(* IEC 61131-3 sources: OpenUnit/plc/src, 8 files *)

(* ---- BMS.st ---- *)
(* BMS - Burner Management System (NFPA 85 style)
   Master fuel trip (MFT) with first-out cause, furnace purge (5 min) with permissives, gas
   fuel train (main gas trip valves / vent: double block and bleed), four burner elevation
   light-off sequences (igniter -> main flame proving -> in service, flame failure trips the
   elevation), light-off time limit, watchdog to the hardwired MFT relay in the field.
   The four elevations A..D are processed in a FOR loop over arrays 1..4: their field I/O is
   copied in at the top and out at the bottom.
   Naming: I_* field inputs, Q_* field outputs, P_<PEER>_* peer status, IO_* bridge signals. *)
PROGRAM BMS_MAIN
(*@IO*)
  VAR
    RT : FB_PLC_RUNTIME;
    T_AIRLOW : FB_TONS;
    T_LVLHH : FB_TONS;
    T_LVLLL : FB_TONS;
    T_FLAMELOSS : FB_TONS;
    T_FUELLOSS : FB_TONS;
    T_BFPLOSS : FB_TONS;
    T_HDRLL : FB_TONS;
    T_HDRHH : FB_TONS;
    T_SUPLOW : FB_TONS;
    dts : REAL;
    init : BOOL;
    (* process values *)
    idRun : BOOL;
    fdRun : BOOL;
    airPct : REAL;
    fp : REAL;
    lvl : REAL;
    hdr : REAL;
    sup : REAL;
    anyFlame : BOOL;
    anyBrnOpen : BOOL;
    nInService : DINT;
    bfpAny : BOOL;
    dehTripped : BOOL;
    dehTripPrev : BOOL;
    mgtvOpen : BOOL;
    (* MFT *)
    c : ARRAY[1..18] OF BOOL;   (* MFT conditions, by first-out cause number *)
    firstOut : DINT;
    mftOn : BOOL;
    cause : DINT;
    fuelWas : BOOL;
    lightoffT : REAL;
    lastFuel : REAL;
    (* purge *)
    ppFans : BOOL;
    ppAir : BOOL;
    ppFuelOff : BOOL;
    ppFurn : BOOL;
    ppDrum : BOOL;
    ppNoTrip : BOOL;
    ready : BOOL;
    purgeActive : BOOL;
    purgeT : REAL;
    purgeComplete : BOOL;
    (* gas train: 0 CLOSED, 1 OPENING, 2 OPEN, 3 TRIPPED *)
    trainState : DINT;
    trainT : REAL;
    trainPerm : BOOL;
    trainCmd : BOOL;
    trainOpen : BOOL;
    (* elevations: state 0 OFF, 1 STARTING, 2 IN SERVICE, 3 STOPPING, 4 FLAME FAIL *)
    x : INT;
    elevPerm : BOOL;
    eState : ARRAY[1..4] OF DINT;
    eT : ARRAY[1..4] OF REAL;
    eIgn : ARRAY[1..4] OF BOOL;
    eBrn : ARRAY[1..4] OF BOOL;
    eLossT : ARRAY[1..4] OF REAL;
    flame : ARRAY[1..4] OF BOOL;
    ignFlame : ARRAY[1..4] OF BOOL;
    brnOpen : ARRAY[1..4] OF BOOL;
    startPb : ARRAY[1..4] OF BOOL;
    stopPb : ARRAY[1..4] OF BOOL;
    fired : BOOL;
  END_VAR
  VAR CONSTANT
    AIR_MCR : REAL := 2247.0;       (* t/h *)
    PURGE_TIME : REAL := 300.0;     (* s *)
    LIGHTOFF_TIME : REAL := 900.0;  (* s *)
    S_OFF : DINT := 0;
    S_STARTING : DINT := 1;
    S_IN_SERVICE : DINT := 2;
    S_STOPPING : DINT := 3;
    S_FAIL : DINT := 4;
    TR_CLOSED : DINT := 0;
    TR_OPENING : DINT := 1;
    TR_OPEN : DINT := 2;
    TR_TRIPPED : DINT := 3;
  END_VAR

  (* ---------------------------------------------------------------- runtime services *)
  RT(SIM_MS := I_SIM_TIME_MS, IC_SEQ := IO_IC_SEQ, IC_ID := IO_IC_ID, IC_SNAP := IO_IC_SNAP, CYCLE_MS := 50.0,
     HEARTBEAT := HEARTBEAT, SCAN_COUNT := SCAN_COUNT, SCAN_MS := SCAN_MS, SIM_DT := SIM_DT,
     IC_APPLIED := IC_APPLIED, IC_ACK := IC_ACK);
  dts := RT.DTS;
  init := RT.IC_INIT;
  HEALTHY := IO_COMM_PLANT AND RT.READY;
  COMM_PLANT := IO_COMM_PLANT OR NOT RT.READY;   (* not reported before the bridge has initialised the PLC *)
  COMM_DEH := IO_COMM_DEH OR RT.GRACE OR NOT RT.READY;

  (* field I/O of the four elevations -> arrays *)
  flame[1] := I_FLAME_A; flame[2] := I_FLAME_B; flame[3] := I_FLAME_C; flame[4] := I_FLAME_D;
  ignFlame[1] := I_IGN_A_FLAME; ignFlame[2] := I_IGN_B_FLAME; ignFlame[3] := I_IGN_C_FLAME; ignFlame[4] := I_IGN_D_FLAME;
  brnOpen[1] := I_BRN_A_OPEN; brnOpen[2] := I_BRN_B_OPEN; brnOpen[3] := I_BRN_C_OPEN; brnOpen[4] := I_BRN_D_OPEN;
  startPb[1] := ELEV_A_START; startPb[2] := ELEV_B_START; startPb[3] := ELEV_C_START; startPb[4] := ELEV_D_START;
  stopPb[1] := ELEV_A_STOP; stopPb[2] := ELEV_B_STOP; stopPb[3] := ELEV_C_STOP; stopPb[4] := ELEV_D_STOP;

  (* ---------------------------------------------------------------- initial condition *)
  (* The firing state follows the plant: a fired boiler is on line with its burning elevations
     in service, otherwise the BMS starts tripped (cause 15, power-up) and needs a purge. *)
  IF init THEN
    fired := I_FLAME_A OR I_FLAME_B OR I_FLAME_C OR I_FLAME_D;
    purgeActive := FALSE;
    purgeT := 0.0;
    purgeComplete := FALSE;
    lightoffT := 0.0;
    dehTripPrev := FALSE;
    IF fired THEN
      mftOn := FALSE;
      cause := 0;
      fuelWas := TRUE;
      trainState := TR_OPEN;
    ELSE
      mftOn := TRUE;
      cause := 15;
      fuelWas := FALSE;
      trainState := TR_TRIPPED;
    END_IF;
    trainT := 0.0;
    FOR x := 1 TO 4 DO
      IF flame[x] THEN eState[x] := S_IN_SERVICE; ELSE eState[x] := S_OFF; END_IF;
      eT[x] := 60.0;
      eIgn[x] := FALSE;
      eBrn[x] := flame[x];
      eLossT[x] := 0.0;
    END_FOR;
    lastFuel := I_FUEL_HEAT;
  END_IF;

  IF RT.READY THEN
    idRun := I_ID_A_RUN OR I_ID_B_RUN;
    fdRun := I_FD_A_RUN OR I_FD_B_RUN;
    airPct := I_AIR_FLOW / AIR_MCR * 100.0;
    fp := MEDIAN3(I_FURN_PRESS_A, I_FURN_PRESS_B, I_FURN_PRESS_C);
    lvl := MEDIAN3(I_DRUM_LVL_A, I_DRUM_LVL_B, I_DRUM_LVL_C);
    hdr := I_GAS_HDR_PRESS;
    sup := I_GAS_SUPPLY_PRESS;
    anyFlame := FALSE;
    anyBrnOpen := FALSE;
    nInService := 0;
    FOR x := 1 TO 4 DO
      anyFlame := anyFlame OR flame[x];
      anyBrnOpen := anyBrnOpen OR brnOpen[x] OR eBrn[x];
      IF eState[x] = S_IN_SERVICE THEN nInService := nInService + 1; END_IF;
    END_FOR;
    bfpAny := I_BFP_A_RUN OR I_BFP_B_RUN OR I_BFP_C_RUN;
    dehTripped := IO_COMM_DEH AND P_DEH_TRIPPED;
    mgtvOpen := I_MGTV_OPEN;

    (* ---------------------------------------------------------------- MFT conditions *)
    T_AIRLOW(IN := airPct < 25.0, PT := 3.0, DTS := dts, INIT := init);
    T_LVLHH(IN := VOTE2OO3(I_DRUM_LVL_A > 250.0, I_DRUM_LVL_B > 250.0, I_DRUM_LVL_C > 250.0), PT := 3.0, DTS := dts, INIT := init);
    T_LVLLL(IN := VOTE2OO3(I_DRUM_LVL_A < -300.0, I_DRUM_LVL_B < -300.0, I_DRUM_LVL_C < -300.0), PT := 3.0, DTS := dts, INIT := init);
    T_FLAMELOSS(IN := anyBrnOpen AND NOT anyFlame, PT := 5.0, DTS := dts, INIT := init);
    T_FUELLOSS(IN := fuelWas AND NOT anyBrnOpen, PT := 2.0, DTS := dts, INIT := init);
    T_BFPLOSS(IN := fuelWas AND NOT bfpAny, PT := 10.0, DTS := dts, INIT := init);
    T_HDRLL(IN := nInService > 0 AND hdr < 120.0, PT := 2.0, DTS := dts, INIT := init);
    T_HDRHH(IN := mgtvOpen AND hdr > 4500.0, PT := 1.0, DTS := dts, INIT := init);
    T_SUPLOW(IN := mgtvOpen AND sup < 12.0, PT := 3.0, DTS := dts, INIT := init);
    c[1] := MFT_PB;                                                              (* manual *)
    c[2] := NOT idRun;                                                           (* both ID fans off *)
    c[3] := NOT fdRun;                                                           (* both FD fans off *)
    c[4] := T_AIRLOW.Q;                                                          (* air flow < 25 % *)
    c[5] := VOTE2OO3(I_FURN_PRESS_A > 20.0, I_FURN_PRESS_B > 20.0, I_FURN_PRESS_C > 20.0);    (* furnace HH *)
    c[6] := VOTE2OO3(I_FURN_PRESS_A < -25.0, I_FURN_PRESS_B < -25.0, I_FURN_PRESS_C < -25.0); (* furnace LL *)
    c[7] := T_LVLHH.Q;                                                           (* drum level HH *)
    c[8] := T_LVLLL.Q;                                                           (* drum level LL *)
    c[9] := T_FLAMELOSS.Q;                                                       (* loss of all flame *)
    c[10] := T_FUELLOSS.Q;                                                       (* loss of all fuel *)
    c[11] := dehTripped AND NOT dehTripPrev AND lastFuel > 0.4 * 1620.0;         (* turbine trip, firing > bypass *)
    c[12] := T_BFPLOSS.Q;                                                        (* all BFPs off *)
    c[13] := NOT mftOn AND NOT fuelWas AND lightoffT > LIGHTOFF_TIME;              (* light-off time expired *)
    c[14] := I_BMS_WD_FAIL;                                                      (* watchdog / field I/O *)
    c[15] := FALSE;                                                              (* power-up: set at initialisation *)
    c[16] := T_HDRLL.Q;                                                          (* gas header LL *)
    c[17] := T_HDRHH.Q;                                                          (* gas header HH *)
    c[18] := T_SUPLOW.Q;                                                         (* gas supply low *)
    dehTripPrev := dehTripped;
    lastFuel := I_FUEL_HEAT;
    IF NOT mftOn THEN
      lightoffT := lightoffT + dts;
      firstOut := FIRST_OUT(C1 := c[1], C2 := c[2], C3 := c[3], C4 := c[4], C5 := c[5], C6 := c[6], C7 := c[7], C8 := c[8], C9 := c[9],
                            C10 := c[10], C11 := c[11], C12 := c[12], C13 := c[13], C14 := c[14], C15 := c[15], C16 := c[16], C17 := c[17],
                            C18 := c[18]);
      IF firstOut > 0 THEN
        (* trip: first-out cause, purge lost, all elevations off *)
        mftOn := TRUE;
        cause := firstOut;
        purgeActive := FALSE;
        purgeT := 0.0;
        purgeComplete := FALSE;
        fuelWas := FALSE;
        FOR x := 1 TO 4 DO
          eState[x] := S_OFF;
          eIgn[x] := FALSE;
          eBrn[x] := FALSE;
        END_FOR;
      END_IF;
    END_IF;

    (* ---------------------------------------------------------------- purge *)
    ppFans := idRun AND fdRun;
    ppAir := airPct >= 25.0 AND airPct <= 40.0;
    ppFuelOff := I_MGTV_CLOSED;
    FOR x := 1 TO 4 DO
      ppFuelOff := ppFuelOff AND NOT brnOpen[x] AND NOT eIgn[x];
    END_FOR;
    ppFurn := ABS(fp) < 5.0;
    ppDrum := lvl > -250.0 AND lvl < 200.0;
    ppNoTrip := NOT (c[2] OR c[3] OR c[5] OR c[6] OR c[7] OR c[8] OR c[14]);
    PP_FANS := ppFans;
    PP_AIR := ppAir;
    PP_FUEL_OFF := ppFuelOff;
    PP_FURN := ppFurn;
    PP_DRUM := ppDrum;
    PP_NO_TRIP := ppNoTrip;
    ready := mftOn AND ppFans AND ppAir AND ppFuelOff AND ppFurn AND ppDrum AND ppNoTrip;
    IF PURGE_START AND ready AND NOT purgeComplete THEN
      purgeActive := TRUE;
      purgeT := 0.0;
      purgeComplete := FALSE;
    END_IF;
    IF purgeActive THEN
      IF NOT ready THEN
        purgeActive := FALSE;
      ELSE
        purgeT := purgeT + dts;
        IF purgeT >= PURGE_TIME THEN
          purgeActive := FALSE;
          purgeT := PURGE_TIME;
          purgeComplete := TRUE;
        END_IF;
      END_IF;
    END_IF;
    IF MFT_RESET AND mftOn AND purgeComplete AND ppNoTrip THEN
      mftOn := FALSE;
      cause := 0;
      purgeActive := FALSE;
      purgeT := 0.0;
      purgeComplete := FALSE;
      lightoffT := 0.0;
      fuelWas := FALSE;
      trainState := TR_CLOSED;
      trainT := 0.0;
    END_IF;

    (* ---------------------------------------------------------------- gas fuel train *)
    trainPerm := NOT mftOn AND sup > 16.0 AND I_MGTV_CLOSED;
    IF GAS_TRAIN_OPEN AND trainPerm AND trainState = TR_CLOSED THEN
      trainState := TR_OPENING;
      trainT := 0.0;
    END_IF;
    IF GAS_TRAIN_CLOSE AND nInService = 0 THEN
      trainState := TR_CLOSED;
      trainT := 0.0;
    END_IF;
    IF mftOn AND trainState <> TR_TRIPPED THEN
      trainState := TR_TRIPPED;
      trainT := 0.0;
    END_IF;
    IF trainState = TR_OPENING THEN
      trainT := trainT + dts;
      IF mgtvOpen THEN
        trainState := TR_OPEN;
      ELSIF trainT > 10.0 THEN
        trainState := TR_CLOSED;
        trainT := 0.0;
      END_IF;
    END_IF;
    trainCmd := trainState = TR_OPENING OR trainState = TR_OPEN;
    Q_MGTV_CMD := trainCmd;
    Q_GAS_VENT_CMD := NOT trainCmd;
    trainOpen := trainState = TR_OPEN AND mgtvOpen AND NOT I_GAS_VENT_OPEN;
    GAS_TRAIN_STATE := trainState;
    GAS_TRAIN_PERM := trainPerm;
    GAS_TRAIN_OPENED := trainOpen;

    (* ---------------------------------------------------------------- burner elevations *)
    elevPerm := NOT mftOn AND trainOpen AND airPct > 25.0 AND hdr > 150.0 AND hdr < 3000.0 AND ABS(fp) < 10.0;
    FOR x := 1 TO 4 DO
      IF startPb[x] AND elevPerm AND (eState[x] = S_OFF OR eState[x] = S_FAIL) THEN
        eState[x] := S_STARTING;
        eT[x] := 0.0;
      END_IF;
      IF stopPb[x] THEN
        IF eState[x] = S_STARTING OR eState[x] = S_IN_SERVICE THEN
          eState[x] := S_STOPPING;
          eT[x] := 0.0;
        ELSIF eState[x] = S_FAIL THEN
          eState[x] := S_OFF;
        END_IF;
      END_IF;
      eT[x] := eT[x] + dts;
      CASE eState[x] OF
        1: (* STARTING: igniter, then main burner valves once the igniter flame is proven *)
          eIgn[x] := TRUE;
          IF eT[x] > 6.0 AND NOT ignFlame[x] THEN
            eState[x] := S_FAIL; eIgn[x] := FALSE; eBrn[x] := FALSE; eT[x] := 0.0;   (* igniter flame not proven *)
          ELSIF ignFlame[x] THEN
            eBrn[x] := TRUE;
          END_IF;
          IF eState[x] = S_STARTING AND eBrn[x] AND flame[x] AND eT[x] > 5.0 THEN
            eState[x] := S_IN_SERVICE;
            eT[x] := 0.0;
          ELSIF eState[x] = S_STARTING AND eT[x] > 15.0 THEN
            eState[x] := S_FAIL; eIgn[x] := FALSE; eBrn[x] := FALSE; eT[x] := 0.0;   (* main flame not proven *)
          END_IF;
        2: (* IN SERVICE: igniter off after 10 s, 2 s loss of flame trips the elevation *)
          eBrn[x] := TRUE;
          eIgn[x] := eT[x] < 10.0;
          IF NOT flame[x] THEN eLossT[x] := MIN(2.0, eLossT[x] + dts); ELSE eLossT[x] := 0.0; END_IF;
          IF NOT flame[x] AND eLossT[x] >= 2.0 THEN
            eState[x] := S_FAIL; eIgn[x] := FALSE; eBrn[x] := FALSE; eT[x] := 0.0;   (* loss of flame *)
          END_IF;
        3: (* STOPPING *)
          eBrn[x] := FALSE;
          eIgn[x] := FALSE;
          IF eT[x] > 3.0 THEN eState[x] := S_OFF; END_IF;
      ELSE
        eBrn[x] := FALSE;
        eIgn[x] := FALSE;
      END_CASE;
      IF eState[x] <> S_IN_SERVICE THEN eLossT[x] := 0.0; END_IF;
      IF mftOn THEN
        eBrn[x] := FALSE;
        eIgn[x] := FALSE;
        IF eState[x] <> S_FAIL THEN eState[x] := S_OFF; END_IF;
      END_IF;
    END_FOR;
    nInService := 0;
    FOR x := 1 TO 4 DO
      IF eState[x] = S_IN_SERVICE THEN nInService := nInService + 1; END_IF;
    END_FOR;
    IF nInService > 0 THEN fuelWas := TRUE; END_IF;

    (* arrays -> field outputs and faceplate status *)
    Q_IGN_A_CMD := eIgn[1]; Q_IGN_B_CMD := eIgn[2]; Q_IGN_C_CMD := eIgn[3]; Q_IGN_D_CMD := eIgn[4];
    Q_BRN_A_CMD := eBrn[1]; Q_BRN_B_CMD := eBrn[2]; Q_BRN_C_CMD := eBrn[3]; Q_BRN_D_CMD := eBrn[4];
    ELEV_A_STATE := eState[1]; ELEV_B_STATE := eState[2]; ELEV_C_STATE := eState[3]; ELEV_D_STATE := eState[4];
    ELEV_A_INSERV := eState[1] = S_IN_SERVICE; ELEV_B_INSERV := eState[2] = S_IN_SERVICE;
    ELEV_C_INSERV := eState[3] = S_IN_SERVICE; ELEV_D_INSERV := eState[4] = S_IN_SERVICE;
    ELEV_A_FAIL := eState[1] = S_FAIL; ELEV_B_FAIL := eState[2] = S_FAIL;
    ELEV_C_FAIL := eState[3] = S_FAIL; ELEV_D_FAIL := eState[4] = S_FAIL;
    ELEV_A_PERM := elevPerm; ELEV_B_PERM := elevPerm; ELEV_C_PERM := elevPerm; ELEV_D_PERM := elevPerm;

    (* ---------------------------------------------------------------- outputs & status *)
    Q_MFT_TRIP := mftOn;
    MFT := mftOn;
    MFT_CAUSE := cause;
    PURGE_READY := ready;
    PURGE_ACTIVE := purgeActive;
    PURGE_COMPLETE := purgeComplete;
    IF purgeComplete THEN PURGE_REMAIN := 0.0; ELSE PURGE_REMAIN := PURGE_TIME - purgeT; END_IF;
    IF mftOn OR fuelWas THEN LIGHTOFF_REMAIN := 0.0; ELSE LIGHTOFF_REMAIN := MAX(0.0, LIGHTOFF_TIME - lightoffT); END_IF;
    FUEL_IN_SERVICE := nInService > 0;
    ELEV_INSERV := nInService;
    IF anyFlame THEN FIREBALL := MIN(100.0, I_FUEL_HEAT / 1620.0 * 110.0); ELSE FIREBALL := 0.0; END_IF;
  END_IF;

  (* watchdog to the hardwired MFT relay: the field trips the boiler if this stops changing *)
  Q_BMS_WD := HEARTBEAT;

  (* operator pulses are consumed in the scan they arrive *)
  MFT_PB := FALSE;
  PURGE_START := FALSE;
  MFT_RESET := FALSE;
  GAS_TRAIN_OPEN := FALSE;
  GAS_TRAIN_CLOSE := FALSE;
  ELEV_A_START := FALSE; ELEV_B_START := FALSE; ELEV_C_START := FALSE; ELEV_D_START := FALSE;
  ELEV_A_STOP := FALSE; ELEV_B_STOP := FALSE; ELEV_C_STOP := FALSE; ELEV_D_STOP := FALSE;
END_PROGRAM

(* ---- BOP.st ---- *)
(* BOP - Balance of Plant / Turbine Auxiliaries
   Circulating water, condenser vacuum, condensate pumps, lube oil / jacking oil / turning
   gear, gland steam, vacuum breaker, hotwell level (condenser make-up).
   Naming: I_* field inputs, Q_* field outputs, P_<PEER>_* peer status, IO_* bridge signals;
   all other located variables are this controller's own Modbus registers (HMI faceplates). *)
PROGRAM BOP_MAIN
(*@IO*)
  VAR
    RT : FB_PLC_RUNTIME;
    CWP_A : FB_MOTOR;
    CWP_B : FB_MOTOR;
    VP_A : FB_MOTOR;
    VP_B : FB_MOTOR;
    CEP_A : FB_MOTOR;
    CEP_B : FB_MOTOR;
    AOP : FB_MOTOR;
    EOP : FB_MOTOR;
    JOP : FB_MOTOR;
    TG : FB_MOTOR;
    GLAND : FB_ONOFF;
    VB : FB_ONOFF;
    HW_DUMP : FB_ONOFF;
    LIC_HW : FB_LOOP;
    CEP_LOWP_TMR : FB_TONS;
    dts : REAL;
    init : BOOL;
    speed : REAL;
    condP : REAL;
    loP : REAL;
    hwLvl : REAL;
    vacPoor : BOOL;
    cepPermit : BOOL;
    cepLowP : BOOL;
    tgPermit : BOOL;
    dehTripped : BOOL;
    tripCwpA : BOOL;
    tripCwpB : BOOL;
    tripVpA : BOOL;
    tripVpB : BOOL;
    tripCepA : BOOL;
    tripCepB : BOOL;
  END_VAR

  (* ---------------------------------------------------------------- runtime services *)
  RT(SIM_MS := I_SIM_TIME_MS, IC_SEQ := IO_IC_SEQ, IC_ID := IO_IC_ID, IC_SNAP := IO_IC_SNAP, CYCLE_MS := 50.0,
     HEARTBEAT := HEARTBEAT, SCAN_COUNT := SCAN_COUNT, SCAN_MS := SCAN_MS, SIM_DT := SIM_DT,
     IC_APPLIED := IC_APPLIED, IC_ACK := IC_ACK);
  dts := RT.DTS;
  init := RT.IC_INIT;
  HEALTHY := IO_COMM_PLANT AND RT.READY;
  COMM_PLANT := IO_COMM_PLANT OR NOT RT.READY;   (* not reported before the bridge has initialised the PLC *)
  COMM_DEH := IO_COMM_DEH OR RT.GRACE OR NOT RT.READY;

  (* ---------------------------------------------------------------- built-in initial condition *)
  IF RT.IC_BUILTIN THEN
    CWP_A_MODE := 1; CWP_B_MODE := 1; VP_A_MODE := 1; VP_B_MODE := 1; CEP_A_MODE := 1; CEP_B_MODE := 1;
    AOP_MODE := 1; EOP_MODE := 1; JOP_MODE := 1; TG_MODE := 1;
    HW_DUMP_MODE := 1;
    LIC_HW_OUT := I_MAKEUP_FB;
    IF IO_IC_ID >= 2 THEN
      LIC_HW_MODE := 1;
    ELSE
      LIC_HW_MODE := 0;
    END_IF;
  END_IF;

  IF RT.READY THEN
    speed := MEDIAN3(I_SPEED_A, I_SPEED_B, I_SPEED_C);
    condP := I_COND_PRESS;
    loP := I_LO_PRESS;
    hwLvl := I_HW_LVL;

    (* Standby pumps start on the latched trip of the duty pump (cleared by the operator's STOP) *)
    tripCwpA := I_CWP_A_TRIP OR (CWP_A.LATCHED AND NOT init);
    tripCwpB := I_CWP_B_TRIP OR (CWP_B.LATCHED AND NOT init);
    tripVpA := I_VP_A_TRIP OR (VP_A.LATCHED AND NOT init);
    tripVpB := I_VP_B_TRIP OR (VP_B.LATCHED AND NOT init);
    tripCepA := I_CEP_A_TRIP OR (CEP_A.LATCHED AND NOT init);
    tripCepB := I_CEP_B_TRIP OR (CEP_B.LATCHED AND NOT init);

    (* ---- circulating water: the standby pump starts when the duty pump trips *)
    CWP_A(RUN_FB := I_CWP_A_RUN, TRIP_FB := I_CWP_A_TRIP, AUTO_START := tripCwpB, SYNC := init,
          START := CWP_A_START, STOP := CWP_A_STOP, MODE := CWP_A_MODE, CMD := Q_CWP_A_CMD,
          RUN := CWP_A_RUN, TRIP := CWP_A_TRIP, PERM := CWP_A_PERM, ILK_T := CWP_A_ILK);
    CWP_B(RUN_FB := I_CWP_B_RUN, TRIP_FB := I_CWP_B_TRIP, AUTO_START := tripCwpA, SYNC := init,
          START := CWP_B_START, STOP := CWP_B_STOP, MODE := CWP_B_MODE, CMD := Q_CWP_B_CMD,
          RUN := CWP_B_RUN, TRIP := CWP_B_TRIP, PERM := CWP_B_PERM, ILK_T := CWP_B_ILK);

    (* ---- vacuum pumps: standby starts on partner trip or poor vacuum *)
    vacPoor := condP > 150.0 AND I_GLAND_ON;
    VP_A(RUN_FB := I_VP_A_RUN, TRIP_FB := I_VP_A_TRIP, AUTO_START := tripVpB OR (vacPoor AND I_VP_B_RUN), SYNC := init,
         START := VP_A_START, STOP := VP_A_STOP, MODE := VP_A_MODE, CMD := Q_VP_A_CMD,
         RUN := VP_A_RUN, TRIP := VP_A_TRIP, PERM := VP_A_PERM, ILK_T := VP_A_ILK);
    VP_B(RUN_FB := I_VP_B_RUN, TRIP_FB := I_VP_B_TRIP, AUTO_START := tripVpA OR (vacPoor AND I_VP_A_RUN), SYNC := init,
         START := VP_B_START, STOP := VP_B_STOP, MODE := VP_B_MODE, CMD := Q_VP_B_CMD,
         RUN := VP_B_RUN, TRIP := VP_B_TRIP, PERM := VP_B_PERM, ILK_T := VP_B_ILK);

    (* ---- condensate pumps: need hotwell level; standby starts on trip or low discharge pressure *)
    cepPermit := hwLvl > 300.0;
    CEP_LOWP_TMR(IN := I_CEP_PRESS < 12.0 AND (I_CEP_A_RUN OR I_CEP_B_RUN), PT := 5.0, DTS := dts, INIT := init);
    cepLowP := CEP_LOWP_TMR.Q;
    CEP_A(RUN_FB := I_CEP_A_RUN, TRIP_FB := I_CEP_A_TRIP, PERMIT := cepPermit, AUTO_START := tripCepB OR (cepLowP AND I_CEP_B_RUN), SYNC := init,
          START := CEP_A_START, STOP := CEP_A_STOP, MODE := CEP_A_MODE, CMD := Q_CEP_A_CMD,
          RUN := CEP_A_RUN, TRIP := CEP_A_TRIP, PERM := CEP_A_PERM, ILK_T := CEP_A_ILK);
    CEP_B(RUN_FB := I_CEP_B_RUN, TRIP_FB := I_CEP_B_TRIP, PERMIT := cepPermit, AUTO_START := tripCepA OR (cepLowP AND I_CEP_A_RUN), SYNC := init,
          START := CEP_B_START, STOP := CEP_B_STOP, MODE := CEP_B_MODE, CMD := Q_CEP_B_CMD,
          RUN := CEP_B_RUN, TRIP := CEP_B_TRIP, PERM := CEP_B_PERM, ILK_T := CEP_B_ILK);

    (* ---- lube oil, jacking oil, turning gear *)
    AOP(RUN_FB := I_AOP_RUN, TRIP_FB := I_AOP_TRIP, AUTO_START := loP < 1.0, SYNC := init,
        START := AOP_START, STOP := AOP_STOP, MODE := AOP_MODE, CMD := Q_AOP_CMD,
        RUN := AOP_RUN, TRIP := AOP_TRIP, PERM := AOP_PERM, ILK_T := AOP_ILK);
    EOP(RUN_FB := I_EOP_RUN, TRIP_FB := I_EOP_TRIP, AUTO_START := loP < 0.7, SYNC := init,
        START := EOP_START, STOP := EOP_STOP, MODE := EOP_MODE, CMD := Q_EOP_CMD,
        RUN := EOP_RUN, TRIP := EOP_TRIP, PERM := EOP_PERM, ILK_T := EOP_ILK);
    JOP(RUN_FB := I_JOP_RUN, TRIP_FB := I_JOP_TRIP, AUTO_START := speed < 600.0 AND loP > 0.5, AUTO_STOP := speed > 700.0, SYNC := init,
        START := JOP_START, STOP := JOP_STOP, MODE := JOP_MODE, CMD := Q_JOP_CMD,
        RUN := JOP_RUN, TRIP := JOP_TRIP, PERM := JOP_PERM, ILK_T := JOP_ILK);
    tgPermit := speed < 5.0 AND I_JOP_RUN AND loP > 1.0;
    TG(RUN_FB := I_TG_RUN, TRIP_FB := I_TG_TRIP, PERMIT := tgPermit OR I_TG_RUN, AUTO_START := tgPermit, ILK := loP < 0.5, SYNC := init,
       START := TG_START, STOP := TG_STOP, MODE := TG_MODE, CMD := Q_TG_CMD,
       RUN := TG_RUN, TRIP := TG_TRIP, PERM := TG_PERM, ILK_T := TG_ILK);

    (* ---- gland steam, vacuum breaker (only with the turbine tripped and below 2400 rpm), hotwell dump *)
    GLAND(OPENED_FB := I_GLAND_ON, SYNC := init,
          OPEN := GLAND_OPEN, CLOSE := GLAND_CLOSE, MODE := GLAND_MODE, CMD := Q_GLAND_CMD,
          OPENED := GLAND_OPENED, CLOSED := GLAND_CLOSED, PERM := GLAND_PERM, ILK := GLAND_ILK);
    IF IO_COMM_DEH THEN
      dehTripped := P_DEH_TRIPPED;
    ELSE
      dehTripped := TRUE;
    END_IF;
    VB(OPENED_FB := I_VB_OPEN, PERMIT := dehTripped AND speed < 2400.0, SYNC := init,
       OPEN := VB_OPEN, CLOSE := VB_CLOSE, MODE := VB_MODE, CMD := Q_VB_CMD,
       OPENED := VB_OPENED, CLOSED := VB_CLOSED, PERM := VB_PERM, ILK := VB_ILK);
    HW_DUMP(OPENED_FB := I_HW_DUMP_OPEN, AUTO_OPEN := hwLvl > 1100.0, AUTO_CLOSE := hwLvl < 900.0, SYNC := init,
            OPEN := HW_DUMP_OPEN, CLOSE := HW_DUMP_CLOSE, MODE := HW_DUMP_MODE, CMD := Q_HW_DUMP_CMD,
            OPENED := HW_DUMP_OPENED, CLOSED := HW_DUMP_CLOSED, PERM := HW_DUMP_PERM, ILK := HW_DUMP_ILK);

    (* ---- hotwell level via condenser make-up *)
    LIC_HW(PV_IN := hwLvl, DTS := dts, RESYNC := RT.RESYNC, PV_MIN := 0.0, PV_MAX := 1500.0,
           SP := LIC_HW_SP, OUT := LIC_HW_OUT, MODE := LIC_HW_MODE, KP := LIC_HW_KP, TI := LIC_HW_TI, TD := LIC_HW_TD,
           PV := LIC_HW_PV, CSP := LIC_HW_CSP, STS := LIC_HW_STS);
    Q_MAKEUP_DMD := LIC_HW.Q;

    VAC_OK := condP < 200.0;
    CW_OK := I_CWP_A_RUN OR I_CWP_B_RUN;
    LO_OK := loP > 1.0;
    COND_PRESS := condP;
  END_IF;
END_PROGRAM

(* ---- CCS.st ---- *)
(* CCS - Unit Coordinated Control
   Unit control modes BASE / BOILER FOLLOW / TURBINE FOLLOW / COORDINATED with permissives
   (a mode whose permissive drops degrades automatically), unit load demand with ramp rate,
   GO / HOLD, frequency bias, capMw limit from the burner elevations in service and fan /
   BFP runbacks, sliding or fixed throttle pressure setpoint, boiler master (PIC_TP) with
   load feed-forward and fast cut-back on load rejection.
   Naming: I_* field inputs, P_<PEER>_* peer status, W_<PEER>_* values written into peers
   (CMB boiler demand, DEH load / pressure references, STC feed-forward), IO_* bridge signals. *)
PROGRAM CCS_MAIN
(*@IO*)
  VAR
    RT : FB_PLC_RUNTIME;
    PIC_TP : FB_LOOP;
    dts : REAL;
    init : BOOL;
    mw : REAL;
    pms : REAL;
    gcb : BOOL;
    gcbPrev : BOOL;
    gcbOpened : BOOL;
    mft : BOOL;
    elevIn : DINT;
    remReady : BOOL;
    latched : BOOL;
    fmAuto : BOOL;
    airAuto : BOOL;
    furnAuto : BOOL;
    rbFan : BOOL;
    lvlAuto : BOOL;
    rbBfp : BOOL;
    bfPerm : BOOL;
    ccPerm : BOOL;
    tfPerm : BOOL;
    req : DINT;
    active : DINT;
    prevActive : DINT;
    dropT : REAL;
    capMw : REAL;
    rbRate : REAL;
    goLatch : BOOL;
    uld : REAL;
    psp : REAL;
    dev : REAL;
    blockInc : BOOL;
    blockDec : BOOL;
    rbActive : BOOL;
    tgt : REAL;
    lim : REAL;
    stepR : REAL;
    d : REAL;
    df : REAL;
    dfDb : REAL;
    fbias : REAL;
    uldF : REAL;
    loadForP : REAL;
    loadPct : REAL;
    pTarget : REAL;
    pr : REAL;
    bmTrk : BOOL;
    bmTrkVal : REAL;
    ffLoad : REAL;
    cutBack : BOOL;
  END_VAR
  VAR CONSTANT
    RATED : REAL := 700.0;        (* MW *)
    ELEV_MW : REAL := 210.0;      (* unit capability per burner elevation in service *)
    M_BASE : DINT := 0;
    M_BF : DINT := 1;
    M_TF : DINT := 2;
    M_CC : DINT := 3;
  END_VAR

  (* ---------------------------------------------------------------- runtime services *)
  RT(SIM_MS := I_SIM_TIME_MS, IC_SEQ := IO_IC_SEQ, IC_ID := IO_IC_ID, IC_SNAP := IO_IC_SNAP, CYCLE_MS := 50.0,
     HEARTBEAT := HEARTBEAT, SCAN_COUNT := SCAN_COUNT, SCAN_MS := SCAN_MS, SIM_DT := SIM_DT,
     IC_APPLIED := IC_APPLIED, IC_ACK := IC_ACK);
  dts := RT.DTS;
  init := RT.IC_INIT;
  HEALTHY := IO_COMM_PLANT AND RT.READY;
  COMM_PLANT := IO_COMM_PLANT OR NOT RT.READY;   (* not reported before the bridge has initialised the PLC *)
  COMM_DEH := IO_COMM_DEH OR RT.GRACE OR NOT RT.READY;
  COMM_CMB := IO_COMM_CMB OR RT.GRACE OR NOT RT.READY;
  COMM_FWC := IO_COMM_FWC OR RT.GRACE OR NOT RT.READY;
  COMM_BMS := IO_COMM_BMS OR RT.GRACE OR NOT RT.READY;
  COMM_STC := IO_COMM_STC OR RT.GRACE OR NOT RT.READY;

  mw := I_GEN_MW;
  pms := I_MS_PRESS;
  gcb := I_GCB_CLOSED;
  IF init THEN
    uld := mw;
    psp := pms;
    goLatch := FALSE;
    dropT := 0.0;
    gcbPrev := FALSE;
    prevActive := MODE_REQ;
  END_IF;

  (* ---------------------------------------------------------------- built-in initial condition *)
  IF RT.IC_BUILTIN THEN
    IF mw > 50.0 THEN ULD_TARGET := mw; ELSE ULD_TARGET := 700.0; END_IF;
    IF IO_IC_ID >= 4 THEN MODE_REQ := M_CC; PIC_TP_MODE := 1; ELSE MODE_REQ := M_BASE; PIC_TP_MODE := 0; END_IF;
    prevActive := MODE_REQ;
    PIC_TP_OUT := I_FUEL_HEAT / 1620.0 * 100.0;
  END_IF;

  IF RT.READY THEN
    (* peer status: the I/O bridge keeps the last good values while a peer is unreachable *)
    mft := P_BMS_MFT;
    elevIn := P_BMS_ELEV_INSERV;
    remReady := P_DEH_REM_READY;
    latched := P_DEH_LATCHED;
    fmAuto := P_CMB_FM_AUTO;
    airAuto := P_CMB_AIR_AUTO;
    furnAuto := P_CMB_FURN_AUTO;
    rbFan := P_CMB_RB_FAN;
    lvlAuto := P_FWC_LVL_AUTO;
    rbBfp := P_FWC_RB_BFP;

    (* ---------------------------------------------------------------- mode management *)
    bfPerm := fmAuto AND airAuto AND furnAuto AND NOT mft AND gcb;
    ccPerm := bfPerm AND remReady AND lvlAuto;
    tfPerm := remReady AND latched AND NOT mft;
    CC_PERM := ccPerm;
    BF_PERM := bfPerm;
    TF_PERM := tfPerm;
    req := MODE_REQ;
    active := req;
    IF NOT RT.GRACE THEN
      IF req = M_CC AND NOT ccPerm THEN
        IF bfPerm THEN active := M_BF; ELSE active := M_BASE; END_IF;
      END_IF;
      IF req = M_TF AND NOT tfPerm THEN active := M_BASE; END_IF;
      IF req = M_BF AND NOT bfPerm THEN active := M_BASE; END_IF;
    END_IF;
    IF active <> req THEN
      (* degrade and make the request follow, so the operator must re-select deliberately *)
      IF prevActive = req THEN dropT := 15.0; END_IF;
      MODE_REQ := active;
    END_IF;
    prevActive := active;
    dropT := MAX(0.0, dropT - dts);
    MODE_DROPPED := dropT > 0.0;
    MODE_ACT := active;

    (* ---------------------------------------------------------------- capMw & runback *)
    capMw := MIN(MAX_LOAD, DINT_TO_REAL(elevIn) * ELEV_MW);
    rbRate := 0.0;
    IF rbFan OR rbBfp THEN
      IF rbFan THEN capMw := MIN(capMw, 350.0); ELSE capMw := MIN(capMw, 385.0); END_IF;
      rbRate := 350.0 / 60.0;
    END_IF;
    CAPACITY := capMw;

    (* ---------------------------------------------------------------- unit load demand *)
    IF GO THEN goLatch := TRUE; END_IF;
    IF HOLD THEN goLatch := FALSE; END_IF;
    dev := psp - pms;
    PRESS_DEV := dev;
    blockInc := active = M_CC AND dev > 10.0;
    blockDec := active = M_CC AND dev < -10.0;
    BLOCK_INC := blockInc;
    BLOCK_DEC := blockDec;
    rbActive := FALSE;
    IF active = M_CC OR active = M_TF THEN
      tgt := LIMIT(MIN_LOAD, ULD_TARGET, MAX_LOAD);
      lim := MIN(tgt, capMw);
      IF uld > capMw + 1.0 THEN
        rbActive := TRUE;
        IF rbRate > 0.0 THEN stepR := rbRate * dts; ELSE stepR := 70.0 / 60.0 * dts; END_IF;
        uld := MAX(capMw, uld - stepR);
        ULD_TARGET := lim;
      ELSIF goLatch THEN
        stepR := ULD_RATE / 60.0 * dts;
        d := LIMIT(-stepR, lim - uld, stepR);
        IF (d > 0.0 AND blockInc) OR (d < 0.0 AND blockDec) THEN d := 0.0; END_IF;
        uld := uld + d;
        IF ABS(lim - uld) < 0.05 THEN goLatch := FALSE; END_IF;
      END_IF;
    ELSE
      uld := MAX(0.0, mw);
      goLatch := FALSE;
    END_IF;
    RB_ACTIVE := rbActive OR ((rbFan OR rbBfp) AND gcb);
    RB_TARGET := capMw;
    RAMPING := goLatch;
    ULD_ACT := uld;
    (* primary frequency response, 5 % droop with 15 mHz deadband, +/- 70 MW *)
    df := I_GRID_FREQ - 60.0;
    dfDb := 0.0;
    IF df > 0.015 THEN dfDb := df - 0.015; ELSIF df < -0.015 THEN dfDb := df + 0.015; END_IF;
    fbias := 0.0;
    IF FREQ_BIAS <> 0 AND active = M_CC THEN
      fbias := LIMIT(-70.0, -dfDb / 60.0 / 0.05 * RATED, 70.0);
    END_IF;
    uldF := uld + fbias;
    ULD_FREQ := uldF;

    (* ---------------------------------------------------------------- pressure setpoint *)
    IF active = M_CC OR active = M_TF THEN loadForP := uld; ELSE loadForP := mw; END_IF;
    IF PRESS_MODE = 1 THEN
      (* sliding pressure: 90 bar below 30 % load, 167 bar above 90 %, linear between *)
      loadPct := loadForP / RATED * 100.0;
      IF loadPct <= 30.0 THEN
        pTarget := 90.0;
      ELSIF loadPct >= 90.0 THEN
        pTarget := 167.0;
      ELSE
        pTarget := 90.0 + (loadPct - 30.0) / 60.0 * 77.0;
      END_IF;
    ELSE
      pTarget := PRESS_FIXED;
    END_IF;
    pr := PRESS_RATE / 60.0 * dts;
    IF active = M_BASE THEN
      psp := pms;
    ELSIF NOT RT.RESYNC THEN
      psp := psp + LIMIT(-pr, pTarget - psp, pr);
    END_IF;
    PRESS_SP := psp;

    (* ---------------------------------------------------------------- boiler master *)
    IF active = M_BF OR active = M_CC THEN PIC_TP_MODE := 1; END_IF;
    PIC_TP_SP := psp;
    bmTrk := FALSE;
    bmTrkVal := 0.0;
    IF mft THEN
      bmTrk := TRUE;
      bmTrkVal := 0.0;
    ELSIF NOT fmAuto THEN
      (* fuel master not in CAS: follow the actual firing so its transfer to CAS is bumpless *)
      bmTrk := TRUE;
      bmTrkVal := I_FUEL_HEAT / 1620.0 * 100.0;
    ELSIF active = M_TF THEN
      bmTrk := TRUE;
      bmTrkVal := uldF / RATED * 100.0 * 1.04;
    END_IF;
    IF active = M_CC THEN ffLoad := uldF; ELSE ffLoad := mw; END_IF;
    (* fast cut-back: on load rejection run the boiler back to what the HP / LP bypass can pass *)
    gcbOpened := NOT gcb AND gcbPrev;
    gcbPrev := gcb;
    cutBack := gcbOpened AND PIC_TP.Q > 40.0 AND NOT mft;
    IF cutBack THEN PIC_TP_OUT := 35.0; END_IF;
    PIC_TP(PV_IN := pms, FF := ffLoad / RATED * 100.0, FORCE_MAN := active = M_BASE OR active = M_TF OR mft,
           TRK := bmTrk, TRK_VAL := bmTrkVal,
           DTS := dts, RESYNC := RT.RESYNC OR cutBack, PV_MIN := 0.0, PV_MAX := 200.0, OUT_MIN := 0.0, OUT_MAX := 110.0, SP_TRACK := FALSE,
           SP := PIC_TP_SP, OUT := PIC_TP_OUT, MODE := PIC_TP_MODE, KP := PIC_TP_KP, TI := PIC_TP_TI, TD := PIC_TP_TD,
           PV := PIC_TP_PV, CSP := PIC_TP_CSP, STS := PIC_TP_STS);
    BLR_DMD := PIC_TP.Q;

    (* ---------------------------------------------------------------- peer outputs *)
    W_CMB_BLR_DMD_REM := PIC_TP.Q;
    IF active = M_BF OR active = M_CC THEN W_CMB_CCS_BM_AUTO := 1; ELSE W_CMB_CCS_BM_AUTO := 0; END_IF;
    W_DEH_LOAD_REF_REM := uld;
    W_DEH_PRESS_SP_REM := psp;
    IF active = M_CC THEN W_DEH_CCS_REQ := 1; ELSIF active = M_TF THEN W_DEH_CCS_REQ := 2; ELSE W_DEH_CCS_REQ := 0; END_IF;
    W_STC_BLR_DMD_FF := PIC_TP.Q;
  END_IF;

  GO := FALSE;
  HOLD := FALSE;
END_PROGRAM

(* ---- CMB.st ---- *)
(* CMB - Combustion & Draft Control
   Fuel master (gas flow -> gas control valve) on the CCS boiler demand with air/fuel
   cross-limiting and elevation capacity limit; total air flow (FD master) with O2 trim and
   minimum (purge) air; furnace pressure (ID master) with FD feed-forward and an MFT kicker;
   fan start permissives and interlocks; fuel runback kicker and fan runback request.
   Naming: I_* field inputs, Q_* field outputs, P_<PEER>_* peer status, IO_* bridge signals.
   BLR_DMD_REM / CCS_BM_AUTO / CCS_HB are written into this PLC by CCS. *)
PROGRAM CMB_MAIN
(*@IO*)
  VAR
    RT : FB_PLC_RUNTIME;
    APH_A : FB_MOTOR;
    APH_B : FB_MOTOR;
    ID_A : FB_MOTOR;
    ID_B : FB_MOTOR;
    FD_A : FB_MOTOR;
    FD_B : FB_MOTOR;
    FIC_GAS : FB_LOOP;
    FIC_AIR : FB_LOOP;
    AIC_O2 : FB_LOOP;
    PIC_FURN : FB_LOOP;
    SC_FDA : FB_STATION;
    SC_FDB : FB_STATION;
    SC_IDA : FB_STATION;
    SC_IDB : FB_STATION;
    T_KICK : FB_TONS;
    dts : REAL;
    init : BOOL;
    keep : BOOL;
    bmsOk : BOOL;
    mft : BOOL;
    elevIn : DINT;
    trainOpen : BOOL;
    aph : BOOL;
    idAny : BOOL;
    fdBoth : BOOL;
    idTripPrevA : BOOL;
    idTripPrevB : BOOL;
    blrLatch : REAL;
    blr : REAL;
    gasFlow : REAL;
    air : REAL;
    capacity : REAL;
    gasByAir : REAL;
    gasRaw : REAL;
    gasDmd : REAL;
    hdr : REAL;
    gfcv : REAL;
    fuelTrk : BOOL;
    fuelTrkVal : REAL;
    fansNow : DINT;
    fansPrev : DINT;
    steamPct : REAL;
    o2Prog : REAL;
    airCas : BOOL;
    airDmd : REAL;
    nFdRun : DINT;
    nFdAuto : DINT;
    fdAvg : REAL;
    fdMaster : REAL;
    fp : REAL;
    kicking : BOOL;
    nIdRun : DINT;
    nIdAuto : DINT;
    idAvg : REAL;
    fdRef : REAL;
    ffFurn : REAL;
    gasLo : REAL;
    gasHi : REAL;
  END_VAR
  VAR CONSTANT
    GAS_LHV : REAL := 49.0;       (* MJ/kg *)
    HEAT_MCR : REAL := 1620.0;       (* MW fuel heat at 100 % boiler demand *)
    GAS_MCR : REAL := 119.0204;   (* t/h at 100 % boiler demand = HEAT_MCR / GAS_LHV * 3.6 *)
    AIR_MCR : REAL := 2247.0;     (* t/h at 100 % boiler demand *)
    STOICH : REAL := 17.15;       (* kg air / kg gas *)
    ELEV_CAP : REAL := 39.3649;   (* t/h per burner elevation in service = 0.3 * GAS_MCR *)
    MCR_STEAM : REAL := 2149.0;
  END_VAR

  (* ---------------------------------------------------------------- runtime services *)
  RT(SIM_MS := I_SIM_TIME_MS, IC_SEQ := IO_IC_SEQ, IC_ID := IO_IC_ID, IC_SNAP := IO_IC_SNAP, CYCLE_MS := 50.0,
     HEARTBEAT := HEARTBEAT, SCAN_COUNT := SCAN_COUNT, SCAN_MS := SCAN_MS, SIM_DT := SIM_DT,
     IC_APPLIED := IC_APPLIED, IC_ACK := IC_ACK);
  dts := RT.DTS;
  init := RT.IC_INIT;
  keep := IO_IC_SNAP;
  HEALTHY := IO_COMM_PLANT AND RT.READY;
  COMM_PLANT := IO_COMM_PLANT OR NOT RT.READY;   (* not reported before the bridge has initialised the PLC *)
  COMM_BMS := IO_COMM_BMS OR RT.GRACE OR NOT RT.READY;
  COMM_CCS := IO_COMM_CCS OR RT.GRACE OR NOT RT.READY;

  IF init THEN
    blrLatch := I_FUEL_HEAT / HEAT_MCR * 100.0;
    idTripPrevA := FALSE;
    idTripPrevB := FALSE;
    fansPrev := -1;
    fdRef := FIC_AIR_OUT;
  END_IF;

  (* ---------------------------------------------------------------- built-in initial condition *)
  IF RT.IC_BUILTIN THEN
    keep := TRUE;   (* fan stations: mode set here, keep their bias *)
    SC_FDA_OUT := I_FD_A_PITCH_FB;
    SC_FDB_OUT := I_FD_B_PITCH_FB;
    SC_IDA_OUT := I_ID_A_VANE_FB;
    SC_IDB_OUT := I_ID_B_VANE_FB;
    IF I_FD_A_RUN THEN SC_FDA_MODE := 1; ELSE SC_FDA_MODE := 0; END_IF;
    IF I_FD_B_RUN THEN SC_FDB_MODE := 1; ELSE SC_FDB_MODE := 0; END_IF;
    IF I_ID_A_RUN THEN SC_IDA_MODE := 1; ELSE SC_IDA_MODE := 0; END_IF;
    IF I_ID_B_RUN THEN SC_IDB_MODE := 1; ELSE SC_IDB_MODE := 0; END_IF;
    FIC_GAS_OUT := I_GFCV_FB;
    FIC_AIR_OUT := (I_FD_A_PITCH_FB + I_FD_B_PITCH_FB) / 2.0;
    PIC_FURN_OUT := (I_ID_A_VANE_FB + I_ID_B_VANE_FB) / 2.0;
    AIC_O2_OUT := 100.0;
    IF IO_IC_ID >= 4 THEN FIC_GAS_MODE := 2; AIC_O2_MODE := 1; ELSE FIC_GAS_MODE := 0; AIC_O2_MODE := 0; END_IF;
    IF IO_IC_ID >= 2 THEN FIC_AIR_MODE := 2; PIC_FURN_MODE := 1; ELSE FIC_AIR_MODE := 0; PIC_FURN_MODE := 0; END_IF;
    fdRef := FIC_AIR_OUT;
  END_IF;

  IF RT.READY THEN
    bmsOk := IO_COMM_BMS;
    IF bmsOk THEN mft := P_BMS_MFT; elevIn := P_BMS_ELEV_INSERV; ELSE mft := TRUE; elevIn := 0; END_IF;
    trainOpen := bmsOk AND P_BMS_GAS_TRAIN_OPENED;

    (* ---- fans: air heaters -> ID fans -> FD fans, vanes / pitch closed to start *)
    aph := I_APH_A_RUN OR I_APH_B_RUN;
    APH_A(RUN_FB := I_APH_A_RUN, TRIP_FB := I_APH_A_TRIP, SYNC := init,
          START := APH_A_START, STOP := APH_A_STOP, MODE := APH_A_MODE, CMD := Q_APH_A_CMD,
          RUN := APH_A_RUN, TRIP := APH_A_TRIP, PERM := APH_A_PERM, ILK_T := APH_A_ILK);
    APH_B(RUN_FB := I_APH_B_RUN, TRIP_FB := I_APH_B_TRIP, SYNC := init,
          START := APH_B_START, STOP := APH_B_STOP, MODE := APH_B_MODE, CMD := Q_APH_B_CMD,
          RUN := APH_B_RUN, TRIP := APH_B_TRIP, PERM := APH_B_PERM, ILK_T := APH_B_ILK);
    ID_A(RUN_FB := I_ID_A_RUN, TRIP_FB := I_ID_A_TRIP, PERMIT := aph AND SC_IDA_OUT <= 5.0, SYNC := init,
         START := ID_A_START, STOP := ID_A_STOP, MODE := ID_A_MODE, CMD := Q_ID_A_CMD,
         RUN := ID_A_RUN, TRIP := ID_A_TRIP, PERM := ID_A_PERM, ILK_T := ID_A_ILK);
    ID_B(RUN_FB := I_ID_B_RUN, TRIP_FB := I_ID_B_TRIP, PERMIT := aph AND SC_IDB_OUT <= 5.0, SYNC := init,
         START := ID_B_START, STOP := ID_B_STOP, MODE := ID_B_MODE, CMD := Q_ID_B_CMD,
         RUN := ID_B_RUN, TRIP := ID_B_TRIP, PERM := ID_B_PERM, ILK_T := ID_B_ILK);
    idAny := I_ID_A_RUN OR I_ID_B_RUN;
    fdBoth := I_FD_A_RUN AND I_FD_B_RUN;
    (* losing an ID fan stops its paired FD fan when both FD fans are running *)
    FD_A(RUN_FB := I_FD_A_RUN, TRIP_FB := I_FD_A_TRIP, PERMIT := idAny AND SC_FDA_OUT <= 5.0, ILK := NOT idAny,
         CMD_SET := I_ID_A_TRIP AND NOT idTripPrevA AND fdBoth, CMD_VAL := FALSE, SYNC := init,
         START := FD_A_START, STOP := FD_A_STOP, MODE := FD_A_MODE, CMD := Q_FD_A_CMD,
         RUN := FD_A_RUN, TRIP := FD_A_TRIP, PERM := FD_A_PERM, ILK_T := FD_A_ILK);
    FD_B(RUN_FB := I_FD_B_RUN, TRIP_FB := I_FD_B_TRIP, PERMIT := idAny AND SC_FDB_OUT <= 5.0, ILK := NOT idAny,
         CMD_SET := I_ID_B_TRIP AND NOT idTripPrevB AND fdBoth, CMD_VAL := FALSE, SYNC := init,
         START := FD_B_START, STOP := FD_B_STOP, MODE := FD_B_MODE, CMD := Q_FD_B_CMD,
         RUN := FD_B_RUN, TRIP := FD_B_TRIP, PERM := FD_B_PERM, ILK_T := FD_B_ILK);
    idTripPrevA := I_ID_A_TRIP;
    idTripPrevB := I_ID_B_TRIP;

    (* ---- boiler demand from the CCS boiler master (held while CCS is not writing) *)
    IF IO_COMM_CCS THEN blrLatch := BLR_DMD_REM; END_IF;
    blr := LIMIT(0.0, blrLatch, 115.0);
    BLR_DMD := blr;

    (* ---- fuel master with cross-limiting *)
    gasFlow := I_GAS_FLOW;
    air := I_AIR_FLOW;
    capacity := DINT_TO_REAL(elevIn) * ELEV_CAP;
    gasByAir := air / (STOICH * 1.07);
    gasRaw := blr / 100.0 * GAS_MCR;
    gasDmd := MAX(0.0, MIN(gasRaw, MIN(gasByAir, capacity)));
    GAS_DMD := gasDmd;
    GAS_CAPACITY := capacity;
    CROSS_LIMIT := elevIn > 0 AND gasRaw > gasByAir + 2.0;
    FUEL_HEAT_EST := gasFlow / 3.6 * GAS_LHV;
    hdr := I_GAS_HDR_PRESS;
    gfcv := I_GFCV_FB;
    fuelTrk := FALSE;
    fuelTrkVal := 0.0;
    IF mft OR NOT trainOpen THEN
      fuelTrk := TRUE;
      fuelTrkVal := 0.0;
    ELSIF elevIn = 0 THEN
      fuelTrk := TRUE;
      fuelTrkVal := LIGHTOFF_POS;
    END_IF;
    (* fuel runback kicker: losing an FD or ID fan at load cuts the gas valve at once *)
    fansNow := 0;
    IF I_FD_A_RUN THEN fansNow := fansNow + 1; END_IF;
    IF I_FD_B_RUN THEN fansNow := fansNow + 1; END_IF;
    IF I_ID_A_RUN THEN fansNow := fansNow + 1; END_IF;
    IF I_ID_B_RUN THEN fansNow := fansNow + 1; END_IF;
    IF fansPrev < 0 THEN fansPrev := fansNow; END_IF;
    IF fansNow < fansPrev AND gasFlow > 0.55 * GAS_MCR AND NOT fuelTrk THEN
      fuelTrk := TRUE;
      fuelTrkVal := FIC_GAS_OUT * 0.6;
    END_IF;
    fansPrev := fansNow;
    IF elevIn > 0 THEN gasLo := MIN_FIRE_POS; ELSE gasLo := 0.0; END_IF;
    IF hdr > 3600.0 THEN gasHi := gfcv; ELSE gasHi := 100.0; END_IF;
    FIC_GAS(PV_IN := gasFlow, CSP_IN := gasDmd, CSP_OK := TRUE, TRK := fuelTrk, TRK_VAL := fuelTrkVal, OUT_LO := gasLo, OUT_HI := gasHi,
            DTS := dts, RESYNC := RT.RESYNC, PV_MIN := 0.0, PV_MAX := 180.0, CAS_CFG := TRUE,
            SP := FIC_GAS_SP, OUT := FIC_GAS_OUT, MODE := FIC_GAS_MODE, KP := FIC_GAS_KP, TI := FIC_GAS_TI, TD := FIC_GAS_TD,
            PV := FIC_GAS_PV, CSP := FIC_GAS_CSP, STS := FIC_GAS_STS);
    Q_GFCV_DMD := FIC_GAS.Q;
    FM_AUTO := FIC_GAS_MODE = 2 AND elevIn > 0;

    (* ---- air flow with O2 trim *)
    steamPct := I_STEAM_FLOW / MCR_STEAM * 100.0;
    o2Prog := FGEN5(X := steamPct, X1 := 0.0, Y1 := 5.0, X2 := 30.0, Y2 := 4.0, X3 := 60.0, Y3 := 2.6, X4 := 100.0, Y4 := 2.0, X5 := 100.0, Y5 := 2.0);
    IF AIC_O2_MODE <> 0 THEN AIC_O2_SP := o2Prog + O2_BIAS; END_IF;
    O2_SP_PROG := o2Prog;
    airCas := FIC_AIR_MODE = 2;
    AIC_O2(PV_IN := I_O2, TRK := mft OR elevIn = 0 OR blr < 20.0 OR NOT airCas, TRK_VAL := 100.0,
           DTS := dts, RESYNC := RT.RESYNC, PV_MIN := 0.0, PV_MAX := 10.0, OUT_MIN := 80.0, OUT_MAX := 120.0, SP_TRACK := FALSE,
           SP := AIC_O2_SP, OUT := AIC_O2_OUT, MODE := AIC_O2_MODE, KP := AIC_O2_KP, TI := AIC_O2_TI, TD := AIC_O2_TD,
           PV := AIC_O2_PV, CSP := AIC_O2_CSP, STS := AIC_O2_STS);
    airDmd := MAX(FGEN5(X := blr, X1 := 0.0, Y1 := 30.0, X2 := 30.0, Y2 := 38.0, X3 := 60.0, Y3 := 64.0, X4 := 100.0, Y4 := 100.0, X5 := 110.0, Y5 := 110.0)
                  / 100.0 * AIR_MCR * (AIC_O2.Q / 100.0),
                  MAX(gasFlow * STOICH * 1.1, PURGE_AIR));
    AIR_DMD := airDmd;
    nFdRun := 0; nFdAuto := 0; fdAvg := 0.0;
    IF I_FD_A_RUN THEN nFdRun := nFdRun + 1; fdAvg := fdAvg + SC_FDA_OUT; IF SC_FDA_MODE = 1 THEN nFdAuto := nFdAuto + 1; END_IF; END_IF;
    IF I_FD_B_RUN THEN nFdRun := nFdRun + 1; fdAvg := fdAvg + SC_FDB_OUT; IF SC_FDB_MODE = 1 THEN nFdAuto := nFdAuto + 1; END_IF; END_IF;
    IF nFdRun > 0 THEN fdAvg := fdAvg / DINT_TO_REAL(nFdRun); END_IF;
    FIC_AIR(PV_IN := air, CSP_IN := airDmd, CSP_OK := TRUE, TRK := nFdAuto = 0, TRK_VAL := fdAvg,
            DTS := dts, RESYNC := RT.RESYNC, PV_MIN := 0.0, PV_MAX := 3200.0, CAS_CFG := TRUE,
            SP := FIC_AIR_SP, OUT := FIC_AIR_OUT, MODE := FIC_AIR_MODE, KP := FIC_AIR_KP, TI := FIC_AIR_TI, TD := FIC_AIR_TD,
            PV := FIC_AIR_PV, CSP := FIC_AIR_CSP, STS := FIC_AIR_STS);
    fdMaster := FIC_AIR.Q;
    SC_FDA(AUTO_IN := fdMaster, FB_IN := I_FD_A_PITCH_FB, FORCE_MAN := NOT I_FD_A_RUN, TRK := NOT I_FD_A_RUN, TRK_VAL := 0.0,
           RATE := 4.0, DTS := dts, INIT := init, INIT_KEEP := keep,
           OUT := SC_FDA_OUT, MODE := SC_FDA_MODE, BIAS := SC_FDA_BIAS, IN_TAG := SC_FDA_IN, FB_TAG := SC_FDA_FB, STS := SC_FDA_STS);
    SC_FDB(AUTO_IN := fdMaster, FB_IN := I_FD_B_PITCH_FB, FORCE_MAN := NOT I_FD_B_RUN, TRK := NOT I_FD_B_RUN, TRK_VAL := 0.0,
           RATE := 4.0, DTS := dts, INIT := init, INIT_KEEP := keep,
           OUT := SC_FDB_OUT, MODE := SC_FDB_MODE, BIAS := SC_FDB_BIAS, IN_TAG := SC_FDB_IN, FB_TAG := SC_FDB_FB, STS := SC_FDB_STS);
    Q_FD_A_PITCH_DMD := SC_FDA.Q;
    Q_FD_B_PITCH_DMD := SC_FDB.Q;
    AIR_AUTO := airCas AND nFdAuto > 0;

    (* ---- furnace pressure (ID master) with FD feed-forward and MFT kicker *)
    fp := MEDIAN3(I_FURN_PRESS_A, I_FURN_PRESS_B, I_FURN_PRESS_C);
    FURN_PRESS_SEL := fp;
    kicking := mft AND T_KICK.ET < 10.0;   (* first 10 s after a master fuel trip *)
    T_KICK(IN := mft, PT := 10.0, DTS := dts, INIT := init);
    nIdRun := 0; nIdAuto := 0; idAvg := 0.0;
    IF I_ID_A_RUN THEN nIdRun := nIdRun + 1; idAvg := idAvg + SC_IDA_OUT; IF SC_IDA_MODE = 1 THEN nIdAuto := nIdAuto + 1; END_IF; END_IF;
    IF I_ID_B_RUN THEN nIdRun := nIdRun + 1; idAvg := idAvg + SC_IDB_OUT; IF SC_IDB_MODE = 1 THEN nIdAuto := nIdAuto + 1; END_IF; END_IF;
    IF nIdRun > 0 THEN idAvg := idAvg / DINT_TO_REAL(nIdRun); END_IF;
    ffFurn := 0.25 * (fdMaster - fdRef);
    IF kicking THEN ffFurn := ffFurn - 12.0; END_IF;
    IF RT.RESYNC OR nIdAuto = 0 THEN fdRef := fdMaster; END_IF;
    fdRef := fdRef + (fdMaster - fdRef) * MIN(1.0, dts / 60.0);
    PIC_FURN(PV_IN := fp, FF := ffFurn, TRK := nIdAuto = 0, TRK_VAL := idAvg,
             DTS := dts, RESYNC := RT.RESYNC, PV_MIN := -15.0, PV_MAX := 15.0, DIRECT := TRUE, SP_TRACK := FALSE,
             SP := PIC_FURN_SP, OUT := PIC_FURN_OUT, MODE := PIC_FURN_MODE, KP := PIC_FURN_KP, TI := PIC_FURN_TI, TD := PIC_FURN_TD,
             PV := PIC_FURN_PV, CSP := PIC_FURN_CSP, STS := PIC_FURN_STS);
    SC_IDA(AUTO_IN := PIC_FURN.Q, FB_IN := I_ID_A_VANE_FB, FORCE_MAN := NOT I_ID_A_RUN, TRK := NOT I_ID_A_RUN, TRK_VAL := 0.0,
           RATE := 6.0, DTS := dts, INIT := init, INIT_KEEP := keep,
           OUT := SC_IDA_OUT, MODE := SC_IDA_MODE, BIAS := SC_IDA_BIAS, IN_TAG := SC_IDA_IN, FB_TAG := SC_IDA_FB, STS := SC_IDA_STS);
    SC_IDB(AUTO_IN := PIC_FURN.Q, FB_IN := I_ID_B_VANE_FB, FORCE_MAN := NOT I_ID_B_RUN, TRK := NOT I_ID_B_RUN, TRK_VAL := 0.0,
           RATE := 6.0, DTS := dts, INIT := init, INIT_KEEP := keep,
           OUT := SC_IDB_OUT, MODE := SC_IDB_MODE, BIAS := SC_IDB_BIAS, IN_TAG := SC_IDB_IN, FB_TAG := SC_IDB_FB, STS := SC_IDB_STS);
    Q_ID_A_VANE_DMD := SC_IDA.Q;
    Q_ID_B_VANE_DMD := SC_IDB.Q;
    FURN_AUTO := PIC_FURN.AUTO AND nIdAuto > 0;

    RB_FAN := (nIdRun < 2 OR nFdRun < 2) AND steamPct > 55.0 AND I_GCB_CLOSED;
  END_IF;
END_PROGRAM

(* ---- DEH.st ---- *)
(* DEH - Turbine Control & Protection (digital electro-hydraulic governor)
   Turbine protection with first-out and latch (reset) permissives; operating modes SPEED
   (run-up through the critical speed bands, synchroniser trim from GEN), LOAD (local load
   reference with frequency droop), REMOTE (load reference from CCS) and PRESSURE (turbine
   follow, throttle pressure from CCS); valve position and throttle pressure limiters; OPC
   (overspeed protection controller) on load rejection; turbine stress evaluator (TSE) limits
   the ramp rates; HP / LP bypass FIXED / FOLLOW pressure control; SH start-up vent.
   Naming: I_* field inputs, Q_* field outputs, P_<PEER>_* peer status, IO_* bridge signals.
   LOAD_REF_REM / PRESS_SP_REM / CCS_REQ are written into this PLC by CCS, SYNC_ADJ /
   SYNC_ACTIVE by GEN. *)
PROGRAM DEH_MAIN
(*@IO*)
  VAR
    RT : FB_PLC_RUNTIME;
    SPD_CTRL : FB_LOOP;
    LOAD_CTRL : FB_LOOP;
    PIC_TPT : FB_LOOP;
    PIC_HPB : FB_LOOP;
    PIC_LPB : FB_LOOP;
    SH_VENT : FB_ONOFF;
    T_VIBHH : FB_TONS;
    T_HPXHH : FB_TONS;
    T_HPBCLOSED : FB_TONS;
    dts : REAL;
    init : BOOL;
    n : REAL;
    gcb : BOOL;
    mw : REAL;
    pms : REAL;
    vib : REAL;
    brg : REAL;
    nOver : INT;
    c : ARRAY[1..12] OF BOOL;   (* trip conditions, by first-out cause number *)
    firstOut : DINT;
    tripActive : BOOL;
    latchPerm : BOOL;
    latch : BOOL;              (* turbine latched (reset) *)
    latchPrev : BOOL;
    latchFell : BOOL;
    spdResync : BOOL;
    cause : DINT;
    req : DINT;
    remoteSel : BOOL;
    dehMode : DINT;            (* 0 TRIPPED, 1 SPEED, 2 LOAD, 3 REMOTE, 4 PRESSURE *)
    gcbPrev : BOOL;
    gcbRose : BOOL;
    gcbFell : BOOL;
    lastMw : REAL;
    opcT : REAL;
    opcLatch : BOOL;
    opc : BOOL;
    hpMetal : REAL;
    flowing : BOOL;
    stressHp : REAL;
    stressIp : REAL;
    stressFactor : REAL;
    spdGo : BOOL;
    loadGo : BOOL;
    spdRef : REAL;
    loadRef : REAL;
    target : REAL;
    rate : REAL;
    banded : BOOL;
    df : REAL;
    dfDb : REAL;
    droopPu : REAL;
    fcorr : REAL;
    tgt : REAL;
    r : REAL;
    tpl : BOOL;
    gvHi : REAL;
    pFilt : REAL;
    gv : REAL;
    spLoad : REAL;
    ffGv : REAL;
    lpbIlk : BOOL;
    follow : BOOL;
    hpbSp : REAL;
    lpbSp : REAL;
    fired : BOOL;
    pd : REAL;
  END_VAR
  VAR CONSTANT
    RPM : REAL := 3600.0;      (* 2-pole generator on a 60 Hz grid *)
    M_TRIPPED : DINT := 0;
    M_SPEED : DINT := 1;
    M_LOAD : DINT := 2;
    M_REMOTE : DINT := 3;
    M_PRESSURE : DINT := 4;
  END_VAR

  (* ---------------------------------------------------------------- runtime services *)
  RT(SIM_MS := I_SIM_TIME_MS, IC_SEQ := IO_IC_SEQ, IC_ID := IO_IC_ID, IC_SNAP := IO_IC_SNAP, CYCLE_MS := 50.0,
     HEARTBEAT := HEARTBEAT, SCAN_COUNT := SCAN_COUNT, SCAN_MS := SCAN_MS, SIM_DT := SIM_DT,
     IC_APPLIED := IC_APPLIED, IC_ACK := IC_ACK);
  dts := RT.DTS;
  init := RT.IC_INIT;
  HEALTHY := IO_COMM_PLANT AND RT.READY;
  COMM_PLANT := IO_COMM_PLANT OR NOT RT.READY;   (* not reported before the bridge has initialised the PLC *)
  COMM_BMS := IO_COMM_BMS OR RT.GRACE OR NOT RT.READY;
  COMM_GEN := IO_COMM_GEN OR RT.GRACE OR NOT RT.READY;
  COMM_CCS := IO_COMM_CCS OR RT.GRACE OR NOT RT.READY;

  n := MEDIAN3(I_SPEED_A, I_SPEED_B, I_SPEED_C);
  gcb := I_GCB_CLOSED;
  mw := I_GEN_MW;
  pms := I_MS_PRESS;

  (* ---------------------------------------------------------------- built-in initial condition *)
  IF RT.IC_BUILTIN THEN
    SH_VENT_MODE := 1;
    SPD_CTRL_MODE := 1; SPD_CTRL_OUT := I_GV_POS;
    LOAD_CTRL_MODE := 1; LOAD_CTRL_OUT := I_GV_POS;
    PIC_TPT_MODE := 1; PIC_TPT_OUT := I_GV_POS;
    PIC_HPB_OUT := I_HPB_POS;
    PIC_LPB_OUT := I_LPB_POS;
    HPB_TARGET := pms;
    IF IO_IC_ID >= 2 THEN PIC_HPB_MODE := 1; PIC_LPB_MODE := 1; ELSE PIC_HPB_MODE := 0; PIC_LPB_MODE := 0; END_IF;
    IF I_MSV_OPEN THEN
      SPD_TARGET := n;
      LOAD_TARGET := mw;
      IF gcb THEN
        MODE_SEL := 1;
        HPB_MODE := 1;
      END_IF;
    END_IF;
  END_IF;

  (* ---------------------------------------------------------------- initial condition: state from the plant *)
  IF init THEN
    latch := I_MSV_OPEN;
    IF latch THEN
      cause := 0;
    ELSIF IO_IC_ID = 1 THEN
      cause := 13;   (* power-up *)
    ELSE
      cause := 0;
    END_IF;
    spdRef := n;
    loadRef := mw;
    spdGo := FALSE;
    loadGo := FALSE;
    opcT := 0.0;
    opcLatch := FALSE;
    IF HPB_MODE = 1 THEN
      hpbSp := pms + 10.0;
      lpbSp := I_HRH_PRESS + 3.0;
    ELSE
      hpbSp := pms;
      lpbSp := MAX(9.0, I_HRH_PRESS);
    END_IF;
    gcbPrev := gcb;
    latchPrev := latch;
    lastMw := mw;
    pFilt := pms;
    gv := I_GV_POS;
  END_IF;

  IF RT.READY THEN
    SPEED := n;

    (* ---------------------------------------------------------------- protection *)
    vib := MAX(MAX(MAX(I_VIB_1, I_VIB_2), MAX(I_VIB_3, I_VIB_4)), MAX(I_VIB_5, I_VIB_6));
    brg := MAX(MAX(MAX(I_BRG_T_1, I_BRG_T_2), MAX(I_BRG_T_3, I_BRG_T_4)), MAX(I_BRG_T_5, I_BRG_T_6));
    MAX_VIB := vib;
    nOver := 0;
    IF I_SPEED_A > RPM * 1.1 THEN nOver := nOver + 1; END_IF;
    IF I_SPEED_B > RPM * 1.1 THEN nOver := nOver + 1; END_IF;
    IF I_SPEED_C > RPM * 1.1 THEN nOver := nOver + 1; END_IF;
    T_VIBHH(IN := vib > 250.0 AND n > 200.0, PT := 2.0, DTS := dts, INIT := init);
    T_HPXHH(IN := I_HP_EXH_TEMP > 450.0, PT := 60.0, DTS := dts, INIT := init);
    c[1] := TRIP_PB;                              (* manual *)
    c[2] := nOver >= 2;                           (* electrical overspeed 110 %, 2 out of 3 *)
    c[3] := I_MECH_OVERSPEED;                     (* mechanical overspeed bolt *)
    c[4] := I_COND_PRESS > 300.0;                 (* low condenser vacuum *)
    c[5] := I_LO_PRESS < 0.6;                     (* low lube oil pressure *)
    c[6] := T_VIBHH.Q;                            (* high shaft vibration *)
    c[7] := ABS(I_AXIAL_DISP) > 1.0;              (* axial displacement *)
    c[8] := T_HPXHH.Q;                            (* HP exhaust temperature *)
    c[9] := IO_COMM_BMS AND P_BMS_MFT;            (* boiler MFT *)
    c[10] := IO_COMM_GEN AND P_GEN_LOCKOUT_86;    (* generator protection 86G *)
    c[11] := brg > 115.0;                         (* bearing temperature *)
    c[12] := I_DEH_WD_FAIL;                       (* watchdog / field I/O *)
    firstOut := FIRST_OUT(C1 := c[1], C2 := c[2], C3 := c[3], C4 := c[4], C5 := c[5], C6 := c[6], C7 := c[7], C8 := c[8], C9 := c[9],
                          C10 := c[10], C11 := c[11], C12 := c[12]);
    IF latch AND firstOut > 0 THEN
      latch := FALSE;
      cause := firstOut;
      spdGo := FALSE;
    END_IF;
    (* a trip condition other than the manual trip blocks the latch *)
    tripActive := c[2] OR c[3] OR c[4] OR c[5] OR c[6] OR c[7] OR c[8] OR c[9] OR c[10] OR c[11] OR c[12];
    latchPerm := NOT latch AND NOT tripActive AND I_COND_PRESS < 200.0 AND I_LO_PRESS > 1.0 AND n < RPM * 1.033 AND NOT gcb;
    LATCH_PERM := latchPerm;
    spdResync := FALSE;
    IF RESET AND latchPerm THEN
      latch := TRUE;
      cause := 0;
      spdRef := n;
      spdGo := FALSE;
      SPD_TARGET := n;
      SPD_CTRL_OUT := 0.0;
      spdResync := TRUE;
    END_IF;
    Q_TURB_TRIP := NOT latch;
    Q_MSV_CMD := latch;
    Q_RSV_CMD := latch;

    (* ---------------------------------------------------------------- mode *)
    IF IO_COMM_CCS THEN req := CCS_REQ; ELSE req := 0; END_IF;
    remoteSel := MODE_SEL = 1;
    dehMode := M_TRIPPED;
    IF latch THEN
      IF NOT gcb THEN
        dehMode := M_SPEED;
      ELSIF remoteSel AND req = 1 THEN
        dehMode := M_REMOTE;
      ELSIF remoteSel AND req = 2 THEN
        dehMode := M_PRESSURE;
      ELSE
        dehMode := M_LOAD;
      END_IF;
    END_IF;
    gcbRose := gcb AND NOT gcbPrev;
    gcbFell := NOT gcb AND gcbPrev;
    gcbPrev := gcb;
    IF gcbRose AND latch THEN
      (* initial load pick-up after synchronising *)
      loadRef := MAX(35.0, mw);
      LOAD_TARGET := MAX(35.0, mw);
      loadGo := FALSE;
    END_IF;
    IF gcbFell AND latch THEN
      (* load rejection: OPC pulse, back to speed control at synchronous speed, and the HP / LP
         bypass holds the boiler at its present pressure *)
      IF lastMw > 210.0 THEN opcT := 3.0; END_IF;
      IF PIC_HPB_MODE <> 0 THEN
        HPB_MODE := 0;
        HPB_TARGET := pms;
        hpbSp := pms;
        lpbSp := MAX(9.0, I_HRH_PRESS);
      END_IF;
      spdRef := RPM;
      SPD_TARGET := RPM;
      spdGo := FALSE;
    END_IF;
    lastMw := mw;

    (* ---------------------------------------------------------------- OPC *)
    opcT := MAX(0.0, opcT - dts);
    IF n > RPM * 1.03 THEN
      opcLatch := TRUE;
    ELSIF n < RPM * 1.01 AND opcT <= 0.0 THEN
      opcLatch := FALSE;
    END_IF;
    opc := latch AND (opcLatch OR opcT > 0.0);
    OPC_ACTIVE := opc;

    (* ---------------------------------------------------------------- turbine stress evaluator *)
    hpMetal := I_HP_METAL_TEMP;
    flowing := I_GV_POS > 1.0 AND I_MSV_OPEN;
    IF flowing THEN
      stressHp := (I_MS_TEMP - 40.0 - hpMetal) / 110.0 * 100.0;
      stressIp := (I_HRH_TEMP - 20.0 - I_IP_METAL_TEMP) / 120.0 * 100.0;
    ELSE
      stressHp := 0.0;
      stressIp := 0.0;
    END_IF;
    STRESS_HP := LIMIT(-100.0, stressHp, 200.0);
    STRESS_IP := LIMIT(-100.0, stressIp, 200.0);
    stressFactor := LIMIT(0.2, (110.0 - MAX(stressHp, stressIp)) / 30.0, 1.0);
    IF hpMetal < 200.0 THEN START_CLASS := 0;
    ELSIF hpMetal < 350.0 THEN START_CLASS := 1;
    ELSIF hpMetal < 450.0 THEN START_CLASS := 2;
    ELSE START_CLASS := 3;
    END_IF;

    (* ---------------------------------------------------------------- speed control *)
    IF GO THEN
      IF dehMode = M_SPEED THEN spdGo := TRUE; ELSE loadGo := TRUE; END_IF;
    END_IF;
    IF HOLD THEN
      spdGo := FALSE;
      loadGo := FALSE;
    END_IF;
    target := LIMIT(0.0, SPD_TARGET, RPM * 1.02);
    IF dehMode = M_SPEED THEN
      rate := SPD_RATE / 60.0 * stressFactor;
      (* critical speed bands 1140-1380, 1860-2100, 2160-2400 rpm: pass at >= 300 rpm/min, never hold *)
      banded := (spdRef > 1140.0 AND spdRef < 1380.0) OR (spdRef > 1860.0 AND spdRef < 2100.0) OR (spdRef > 2160.0 AND spdRef < 2400.0);
      IF banded THEN
        rate := MAX(rate, 300.0 / 60.0);
        IF NOT spdGo AND ABS(target - spdRef) > 1.0 THEN spdGo := TRUE; END_IF;
      END_IF;
      IF spdGo THEN
        spdRef := spdRef + LIMIT(-rate * dts, target - spdRef, rate * dts);
        IF ABS(target - spdRef) < 0.5 THEN spdGo := FALSE; END_IF;
      END_IF;
      IF IO_COMM_GEN AND SYNC_ACTIVE <> 0 AND spdRef >= RPM * 0.983 THEN
        spdRef := LIMIT(RPM * 0.983, spdRef + SYNC_ADJ * dts, RPM * 1.02);
        SPD_TARGET := spdRef;
      END_IF;
    ELSE
      spdRef := n;
      spdGo := FALSE;
    END_IF;
    CRIT_ZONE := dehMode = M_SPEED AND ((n > 1140.0 AND n < 1380.0) OR (n > 1860.0 AND n < 2100.0) OR (n > 2160.0 AND n < 2400.0));
    SPEED_REF := spdRef;
    RAMP_ACTIVE := spdGo OR loadGo;

    (* ---------------------------------------------------------------- load / pressure control *)
    df := I_GRID_FREQ - 60.0;
    dfDb := 0.0;
    IF df > 0.015 THEN dfDb := df - 0.015; ELSIF df < -0.015 THEN dfDb := df + 0.015; END_IF;
    droopPu := MAX(1.0, DROOP) / 100.0;
    fcorr := 0.0;
    IF FREQ_ON <> 0 AND gcb THEN
      fcorr := LIMIT(-70.0, -dfDb / 60.0 / droopPu * 700.0, 70.0);
    END_IF;
    FREQ_CORR := fcorr;
    IF dehMode = M_REMOTE THEN
      loadRef := LOAD_REF_REM;
      LOAD_TARGET := loadRef;
    ELSIF dehMode = M_LOAD THEN
      tgt := LIMIT(0.0, LOAD_TARGET, 720.0);
      IF loadGo THEN
        r := LOAD_RATE / 60.0 * stressFactor * dts;
        loadRef := loadRef + LIMIT(-r, tgt - loadRef, r);
        IF ABS(tgt - loadRef) < 0.05 THEN loadGo := FALSE; END_IF;
      END_IF;
    ELSIF dehMode <> M_PRESSURE THEN
      loadRef := MAX(0.0, mw);
      loadGo := FALSE;
    ELSE
      loadRef := mw;
    END_IF;
    LOAD_REF := loadRef;

    (* throttle pressure limiter and valve position limit *)
    tpl := (dehMode = M_LOAD OR dehMode = M_REMOTE) AND pms < TPL_SP;
    TPL_ACTIVE := tpl;
    gvHi := VPL;
    IF tpl THEN gvHi := MIN(gvHi, MAX(0.0, I_GV_POS - 0.5)); END_IF;
    pFilt := pFilt + (pms - pFilt) * MIN(1.0, dts / 30.0);

    IF NOT latch OR opc THEN
      (* tripped / OPC: all governors track a closed valve *)
      SPD_CTRL(PV_IN := n, TRK := TRUE, TRK_VAL := 0.0, OUT_HI := 1.0E30, FF := 0.0,
               DTS := dts, RESYNC := RT.RESYNC OR spdResync, PV_MIN := 0.0, PV_MAX := 4320.0, SP_TRACK := FALSE,
               SP := SPD_CTRL_SP, OUT := SPD_CTRL_OUT, MODE := SPD_CTRL_MODE, KP := SPD_CTRL_KP, TI := SPD_CTRL_TI, TD := SPD_CTRL_TD,
               PV := SPD_CTRL_PV, CSP := SPD_CTRL_CSP, STS := SPD_CTRL_STS);
      LOAD_CTRL(PV_IN := mw, TRK := TRUE, TRK_VAL := 0.0, OUT_HI := 1.0E30, FF := 0.0,
                DTS := dts, RESYNC := RT.RESYNC, PV_MIN := 0.0, PV_MAX := 800.0, SP_TRACK := FALSE,
                SP := LOAD_CTRL_SP, OUT := LOAD_CTRL_OUT, MODE := LOAD_CTRL_MODE, KP := LOAD_CTRL_KP, TI := LOAD_CTRL_TI, TD := LOAD_CTRL_TD,
                PV := LOAD_CTRL_PV, CSP := LOAD_CTRL_CSP, STS := LOAD_CTRL_STS);
      PIC_TPT(PV_IN := pms, TRK := TRUE, TRK_VAL := 0.0, OUT_HI := 1.0E30,
              DTS := dts, RESYNC := RT.RESYNC, PV_MIN := 0.0, PV_MAX := 200.0, DIRECT := TRUE, SP_TRACK := FALSE,
              SP := PIC_TPT_SP, OUT := PIC_TPT_OUT, MODE := PIC_TPT_MODE, KP := PIC_TPT_KP, TI := PIC_TPT_TI, TD := PIC_TPT_TD,
              PV := PIC_TPT_PV, CSP := PIC_TPT_CSP, STS := PIC_TPT_STS);
      gv := 0.0;
    ELSIF dehMode = M_SPEED THEN
      SPD_CTRL_SP := spdRef;
      SPD_CTRL(PV_IN := n, TRK := FALSE, OUT_HI := gvHi, FF := 0.0,
               DTS := dts, RESYNC := RT.RESYNC OR spdResync, PV_MIN := 0.0, PV_MAX := 4320.0, SP_TRACK := FALSE,
               SP := SPD_CTRL_SP, OUT := SPD_CTRL_OUT, MODE := SPD_CTRL_MODE, KP := SPD_CTRL_KP, TI := SPD_CTRL_TI, TD := SPD_CTRL_TD,
               PV := SPD_CTRL_PV, CSP := SPD_CTRL_CSP, STS := SPD_CTRL_STS);
      gv := SPD_CTRL.Q;
      LOAD_CTRL(PV_IN := mw, TRK := TRUE, TRK_VAL := gv, OUT_HI := 1.0E30, FF := 0.0,
                DTS := dts, RESYNC := RT.RESYNC, PV_MIN := 0.0, PV_MAX := 800.0, SP_TRACK := FALSE,
                SP := LOAD_CTRL_SP, OUT := LOAD_CTRL_OUT, MODE := LOAD_CTRL_MODE, KP := LOAD_CTRL_KP, TI := LOAD_CTRL_TI, TD := LOAD_CTRL_TD,
                PV := LOAD_CTRL_PV, CSP := LOAD_CTRL_CSP, STS := LOAD_CTRL_STS);
      PIC_TPT(PV_IN := pms, TRK := TRUE, TRK_VAL := gv, OUT_HI := 1.0E30,
              DTS := dts, RESYNC := RT.RESYNC, PV_MIN := 0.0, PV_MAX := 200.0, DIRECT := TRUE, SP_TRACK := FALSE,
              SP := PIC_TPT_SP, OUT := PIC_TPT_OUT, MODE := PIC_TPT_MODE, KP := PIC_TPT_KP, TI := PIC_TPT_TI, TD := PIC_TPT_TD,
              PV := PIC_TPT_PV, CSP := PIC_TPT_CSP, STS := PIC_TPT_STS);
    ELSIF dehMode = M_PRESSURE THEN
      PIC_TPT_SP := PRESS_SP_REM;
      PIC_TPT(PV_IN := pms, TRK := FALSE, OUT_HI := gvHi,
              DTS := dts, RESYNC := RT.RESYNC, PV_MIN := 0.0, PV_MAX := 200.0, DIRECT := TRUE, SP_TRACK := FALSE,
              SP := PIC_TPT_SP, OUT := PIC_TPT_OUT, MODE := PIC_TPT_MODE, KP := PIC_TPT_KP, TI := PIC_TPT_TI, TD := PIC_TPT_TD,
              PV := PIC_TPT_PV, CSP := PIC_TPT_CSP, STS := PIC_TPT_STS);
      gv := PIC_TPT.Q;
      SPD_CTRL(PV_IN := n, TRK := TRUE, TRK_VAL := gv, OUT_HI := 1.0E30, FF := 0.0,
               DTS := dts, RESYNC := RT.RESYNC OR spdResync, PV_MIN := 0.0, PV_MAX := 4320.0, SP_TRACK := FALSE,
               SP := SPD_CTRL_SP, OUT := SPD_CTRL_OUT, MODE := SPD_CTRL_MODE, KP := SPD_CTRL_KP, TI := SPD_CTRL_TI, TD := SPD_CTRL_TD,
               PV := SPD_CTRL_PV, CSP := SPD_CTRL_CSP, STS := SPD_CTRL_STS);
      LOAD_CTRL(PV_IN := mw, TRK := TRUE, TRK_VAL := gv, OUT_HI := 1.0E30, FF := 0.0,
                DTS := dts, RESYNC := RT.RESYNC, PV_MIN := 0.0, PV_MAX := 800.0, SP_TRACK := FALSE,
                SP := LOAD_CTRL_SP, OUT := LOAD_CTRL_OUT, MODE := LOAD_CTRL_MODE, KP := LOAD_CTRL_KP, TI := LOAD_CTRL_TI, TD := LOAD_CTRL_TD,
                PV := LOAD_CTRL_PV, CSP := LOAD_CTRL_CSP, STS := LOAD_CTRL_STS);
    ELSE
      (* LOAD / REMOTE: load controller with a valve-area feed-forward at the filtered throttle pressure *)
      spLoad := loadRef + fcorr;
      LOAD_CTRL_SP := spLoad;
      ffGv := LIMIT(0.0, spLoad / 700.0 * 90.0 * (168.0 / MAX(20.0, pFilt + 1.0)), 100.0);
      LOAD_CTRL(PV_IN := mw, TRK := FALSE, OUT_HI := gvHi, FF := ffGv,
                DTS := dts, RESYNC := RT.RESYNC, PV_MIN := 0.0, PV_MAX := 800.0, SP_TRACK := FALSE,
                SP := LOAD_CTRL_SP, OUT := LOAD_CTRL_OUT, MODE := LOAD_CTRL_MODE, KP := LOAD_CTRL_KP, TI := LOAD_CTRL_TI, TD := LOAD_CTRL_TD,
                PV := LOAD_CTRL_PV, CSP := LOAD_CTRL_CSP, STS := LOAD_CTRL_STS);
      gv := LOAD_CTRL.Q;
      SPD_CTRL(PV_IN := n, TRK := TRUE, TRK_VAL := gv, OUT_HI := 1.0E30, FF := 0.0,
               DTS := dts, RESYNC := RT.RESYNC OR spdResync, PV_MIN := 0.0, PV_MAX := 4320.0, SP_TRACK := FALSE,
               SP := SPD_CTRL_SP, OUT := SPD_CTRL_OUT, MODE := SPD_CTRL_MODE, KP := SPD_CTRL_KP, TI := SPD_CTRL_TI, TD := SPD_CTRL_TD,
               PV := SPD_CTRL_PV, CSP := SPD_CTRL_CSP, STS := SPD_CTRL_STS);
      PIC_TPT(PV_IN := pms, TRK := TRUE, TRK_VAL := gv, OUT_HI := 1.0E30,
              DTS := dts, RESYNC := RT.RESYNC, PV_MIN := 0.0, PV_MAX := 200.0, DIRECT := TRUE, SP_TRACK := FALSE,
              SP := PIC_TPT_SP, OUT := PIC_TPT_OUT, MODE := PIC_TPT_MODE, KP := PIC_TPT_KP, TI := PIC_TPT_TI, TD := PIC_TPT_TD,
              PV := PIC_TPT_PV, CSP := PIC_TPT_CSP, STS := PIC_TPT_STS);
    END_IF;
    GV_DEMAND := gv;
    Q_GV_DMD := gv;
    (* valve management: the intercept valves share the flow demand at low load so the reheater
       (held up by the LP bypass) cannot over-drive the IP turbine; fully open above ~67 % *)
    IF latch AND NOT opc THEN Q_ICV_DMD := LIMIT(0.0, gv * 1.5, 100.0); ELSE Q_ICV_DMD := 0.0; END_IF;

    (* ---------------------------------------------------------------- HP / LP bypass *)
    lpbIlk := I_COND_PRESS > 300.0 OR I_CW_FLOW < 15000.0;
    LPB_ILK := lpbIlk;
    latchFell := NOT latch AND latchPrev;
    latchPrev := latch;
    IF latchFell AND PIC_HPB_MODE <> 0 THEN
      (* turbine trip: hold the boiler at its present pressure through the bypass *)
      HPB_MODE := 0;
      HPB_TARGET := pms;
      hpbSp := pms;
      lpbSp := MAX(9.0, I_HRH_PRESS);
    END_IF;
    T_HPBCLOSED(IN := gcb AND I_HPB_POS < 2.0 AND mw > 50.0, PT := 30.0, DTS := dts, INIT := init);
    IF T_HPBCLOSED.Q AND HPB_MODE = 0 THEN HPB_MODE := 1; END_IF;
    follow := HPB_MODE = 1;
    IF follow THEN
      (* FOLLOW: setpoints a margin above the actual pressures, rising slowly, falling at once *)
      tgt := pms + 10.0;
      IF tgt < hpbSp THEN hpbSp := tgt; ELSE hpbSp := MIN(tgt, hpbSp + 5.0 / 60.0 * dts); END_IF;
      tgt := I_HRH_PRESS + 3.0;
      IF tgt < lpbSp THEN lpbSp := tgt; ELSE lpbSp := MIN(tgt, lpbSp + 3.0 / 60.0 * dts); END_IF;
    ELSE
      (* FIXED: ramp to the operator target *)
      r := HPB_RAMP / 60.0 * dts;
      hpbSp := hpbSp + LIMIT(-r, HPB_TARGET - hpbSp, r);
      IF PIC_LPB_MODE <> 0 AND NOT gcb THEN lpbSp := 9.0; END_IF;
    END_IF;
    IF PIC_HPB_MODE <> 0 THEN PIC_HPB_SP := hpbSp; ELSE hpbSp := pms; END_IF;
    IF PIC_LPB_MODE <> 0 THEN PIC_LPB_SP := lpbSp; END_IF;
    PIC_HPB(PV_IN := pms, TRK := lpbIlk, TRK_VAL := 0.0,
            DTS := dts, RESYNC := RT.RESYNC, PV_MIN := 0.0, PV_MAX := 200.0, DIRECT := TRUE, SP_TRACK := FALSE,
            SP := PIC_HPB_SP, OUT := PIC_HPB_OUT, MODE := PIC_HPB_MODE, KP := PIC_HPB_KP, TI := PIC_HPB_TI, TD := PIC_HPB_TD,
            PV := PIC_HPB_PV, CSP := PIC_HPB_CSP, STS := PIC_HPB_STS);
    Q_HPB_DMD := PIC_HPB.Q;
    PIC_LPB(PV_IN := I_HRH_PRESS, TRK := lpbIlk, TRK_VAL := 0.0,
            DTS := dts, RESYNC := RT.RESYNC, PV_MIN := 0.0, PV_MAX := 50.0, DIRECT := TRUE, SP_TRACK := FALSE,
            SP := PIC_LPB_SP, OUT := PIC_LPB_OUT, MODE := PIC_LPB_MODE, KP := PIC_LPB_KP, TI := PIC_LPB_TI, TD := PIC_LPB_TD,
            PV := PIC_LPB_PV, CSP := PIC_LPB_CSP, STS := PIC_LPB_STS);
    Q_LPB_DMD := PIC_LPB.Q;

    (* SH start-up vent: open while raising pressure from cold, closed above 5 bar *)
    fired := IO_COMM_BMS AND P_BMS_FUEL_IN_SERVICE;
    pd := I_DRUM_PRESS;
    SH_VENT(OPENED_FB := I_SH_VENT_OPEN, AUTO_OPEN := fired AND pd < 3.0, AUTO_CLOSE := pd > 5.0, SYNC := init,
            OPEN := SH_VENT_OPEN, CLOSE := SH_VENT_CLOSE, MODE := SH_VENT_MODE, CMD := Q_SH_VENT_CMD,
            OPENED := SH_VENT_OPENED, CLOSED := SH_VENT_CLOSED, PERM := SH_VENT_PERM, ILK := SH_VENT_ILK);

    (* ---------------------------------------------------------------- status *)
    TRIPPED := NOT latch;
    LATCHED := latch;
    MODE := dehMode;
    TRIP_CAUSE := cause;
    AT_SPEED := dehMode = M_SPEED AND ABS(n - RPM) < 18.0;
    REM_READY := latch AND gcb AND remoteSel;
  END_IF;

  (* watchdog to the hardwired turbine trip: the field trips the turbine if this stops changing *)
  Q_DEH_WD := HEARTBEAT;

  RESET := FALSE;
  TRIP_PB := FALSE;
  GO := FALSE;
  HOLD := FALSE;
END_PROGRAM

(* ---- FWC.st ---- *)
(* FWC - Feedwater & Condensate Control
   Drum level: 1-element (level -> FW valve) at low load, 3-element (level master trims a steam
   flow feed-forward, FW flow slave) above 25 % steam flow, bumpless transfer between them.
   Boiler feed pumps: valve differential pressure master (PIC_FWDP) -> speed stations, standby
   pump auto start on a partner trip (it joins the master demand), runback request if fewer than
   two pumps run above 58 % load.  Deaerator level and pegging steam, blowdown, HP heaters.
   Naming: I_* field inputs, Q_* field outputs, P_<PEER>_* peer status, IO_* bridge signals. *)
PROGRAM FWC_MAIN
(*@IO*)
  VAR
    RT : FB_PLC_RUNTIME;
    BFP_A : FB_MOTOR;
    BFP_B : FB_MOTOR;
    BFP_C : FB_MOTOR;
    EBD : FB_ONOFF;
    HPH : FB_ONOFF;
    LIC_DRUM : FB_LOOP;
    FIC_FW : FB_LOOP;
    PIC_FWDP : FB_LOOP;
    SC_BFPA : FB_STATION;
    SC_BFPB : FB_STATION;
    SC_BFPC : FB_STATION;
    LIC_DA : FB_LOOP;
    PIC_DA : FB_LOOP;
    HIC_CBD : FB_STATION;
    T_LTDEV : FB_TONS;
    T_RBBFP : FB_TONS;
    dts : REAL;
    init : BOOL;
    keep : BOOL;
    keepCbd : BOOL;
    lvl : REAL;
    steam : REAL;
    spray : REAL;
    fw : REAL;
    ff : REAL;
    steamPct : REAL;
    e3 : BOOL;
    e3Latch : BOOL;
    e3Changed : BOOL;
    e3Trk : REAL;
    ficCas : BOOL;
    nRun : DINT;
    daLvl : REAL;
    dp : REAL;
    dpSp : REAL;
    anyAuto : BOOL;
    avgScoop : REAL;
    master : REAL;
    tripA : BOOL;
    tripB : BOOL;
    tripC : BOOL;
    runPrevA : BOOL;
    runPrevB : BOOL;
    runPrevC : BOOL;
    joinA : BOOL;
    joinB : BOOL;
    joinC : BOOL;
    cep : BOOL;
  END_VAR
  VAR CONSTANT
    MCR_STEAM : REAL := 2149.0;   (* t/h *)
    TRIM_GAIN : REAL := 12.0;     (* t/h per % of level master output in 3-element mode *)
  END_VAR

  (* ---------------------------------------------------------------- runtime services *)
  RT(SIM_MS := I_SIM_TIME_MS, IC_SEQ := IO_IC_SEQ, IC_ID := IO_IC_ID, IC_SNAP := IO_IC_SNAP, CYCLE_MS := 50.0,
     HEARTBEAT := HEARTBEAT, SCAN_COUNT := SCAN_COUNT, SCAN_MS := SCAN_MS, SIM_DT := SIM_DT,
     IC_APPLIED := IC_APPLIED, IC_ACK := IC_ACK);
  dts := RT.DTS;
  init := RT.IC_INIT;
  keep := IO_IC_SNAP;
  keepCbd := IO_IC_SNAP;
  HEALTHY := IO_COMM_PLANT AND RT.READY;
  COMM_PLANT := IO_COMM_PLANT OR NOT RT.READY;   (* not reported before the bridge has initialised the PLC *)
  COMM_BMS := IO_COMM_BMS OR RT.GRACE OR NOT RT.READY;
  COMM_DEH := IO_COMM_DEH OR RT.GRACE OR NOT RT.READY;

  steam := I_STEAM_FLOW;
  spray := I_SH_SPRAY_FLOW;
  fw := I_FW_FLOW;
  ff := MAX(0.0, steam - spray);
  steamPct := steam / MCR_STEAM * 100.0;
  e3Trk := LIMIT(0.0, 50.0 + (fw - ff) / TRIM_GAIN, 100.0);   (* level master output for a bumpless 3-element start *)

  IF init THEN
    (* element selection as it stands, so the IC does not cause a transfer *)
    IF ELEM_SEL = 1 THEN e3Latch := FALSE; ELSIF ELEM_SEL = 2 THEN e3Latch := TRUE; ELSE e3Latch := steamPct > 25.0; END_IF;
    runPrevA := FALSE; runPrevB := FALSE; runPrevC := FALSE;
    joinA := FALSE; joinB := FALSE; joinC := FALSE;
  END_IF;

  (* ---------------------------------------------------------------- built-in initial condition *)
  IF RT.IC_BUILTIN THEN
    keep := TRUE;   (* BFP stations below are set explicitly *)
    EBD_MODE := 1;
    IF I_BFP_A_RUN THEN BFP_A_MODE := 0; SC_BFPA_OUT := LIMIT(0.0, (I_BFP_A_SPEED - 1500.0) / 39.0, 100.0); ELSE BFP_A_MODE := 1; SC_BFPA_OUT := 0.0; END_IF;
    IF I_BFP_B_RUN THEN BFP_B_MODE := 0; SC_BFPB_OUT := LIMIT(0.0, (I_BFP_B_SPEED - 1500.0) / 39.0, 100.0); ELSE BFP_B_MODE := 1; SC_BFPB_OUT := 0.0; END_IF;
    IF I_BFP_C_RUN THEN BFP_C_MODE := 0; SC_BFPC_OUT := LIMIT(0.0, (I_BFP_C_SPEED - 1500.0) / 39.0, 100.0); ELSE BFP_C_MODE := 1; SC_BFPC_OUT := 0.0; END_IF;
    IF I_BFP_A_RUN AND IO_IC_ID >= 2 THEN SC_BFPA_MODE := 1; ELSE SC_BFPA_MODE := 0; END_IF;
    IF I_BFP_B_RUN AND IO_IC_ID >= 2 THEN SC_BFPB_MODE := 1; ELSE SC_BFPB_MODE := 0; END_IF;
    IF I_BFP_C_RUN AND IO_IC_ID >= 2 THEN SC_BFPC_MODE := 1; ELSE SC_BFPC_MODE := 0; END_IF;
    IF I_BFP_A_RUN THEN PIC_FWDP_OUT := SC_BFPA_OUT;
    ELSIF I_BFP_B_RUN THEN PIC_FWDP_OUT := SC_BFPB_OUT;
    ELSIF I_BFP_C_RUN THEN PIC_FWDP_OUT := SC_BFPC_OUT;
    ELSE PIC_FWDP_OUT := 0.0;
    END_IF;
    FIC_FW_OUT := I_FCV_FB;
    LIC_DA_OUT := I_DA_CV_FB;
    PIC_DA_OUT := I_PEG_FB;
    e3Latch := steamPct > 25.0;
    IF e3Latch THEN LIC_DRUM_OUT := e3Trk; ELSE LIC_DRUM_OUT := I_FCV_FB; END_IF;
    IF IO_IC_ID >= 2 THEN
      LIC_DRUM_MODE := 1; FIC_FW_MODE := 2; PIC_FWDP_MODE := 2; LIC_DA_MODE := 1; PIC_DA_MODE := 1;
    ELSE
      LIC_DRUM_MODE := 0; FIC_FW_MODE := 0; PIC_FWDP_MODE := 0; LIC_DA_MODE := 0; PIC_DA_MODE := 0;
    END_IF;
  END_IF;

  IF RT.READY THEN
    lvl := MEDIAN3(I_DRUM_LVL_A, I_DRUM_LVL_B, I_DRUM_LVL_C);
    DRUM_LVL_SEL := lvl;
    T_LTDEV(IN := ABS(I_DRUM_LVL_A - lvl) > 50.0 OR ABS(I_DRUM_LVL_B - lvl) > 50.0 OR ABS(I_DRUM_LVL_C - lvl) > 50.0,
            PT := 5.0, DTS := dts, INIT := init);
    LT_DEVIATION := T_LTDEV.Q;
    STEAM_FLOW_PCT := steamPct;

    (* ---- drum level: 1-element / 3-element with bumpless transfer *)
    IF ELEM_SEL = 1 THEN
      e3 := FALSE;
    ELSIF ELEM_SEL = 2 THEN
      e3 := TRUE;
    ELSIF e3Latch THEN
      e3 := steamPct > 20.0;
    ELSE
      e3 := steamPct > 25.0;
    END_IF;
    e3Changed := e3 <> e3Latch;
    IF e3Changed THEN
      e3Latch := e3;
      IF e3 THEN LIC_DRUM_OUT := e3Trk; ELSE LIC_DRUM_OUT := I_FCV_FB; END_IF;
    END_IF;
    E3_ACTIVE := e3;
    ficCas := FIC_FW_MODE = 2;
    IF NOT e3 THEN
      (* 1-element: the level controller positions the valve through the flow loop *)
      LIC_DRUM(PV_IN := lvl, TRK := NOT ficCas, TRK_VAL := I_FCV_FB,
               DTS := dts, RESYNC := RT.RESYNC OR e3Changed, PV_MIN := -500.0, PV_MAX := 500.0,
               SP := LIC_DRUM_SP, OUT := LIC_DRUM_OUT, MODE := LIC_DRUM_MODE, KP := LIC_DRUM_KP, TI := LIC_DRUM_TI, TD := LIC_DRUM_TD,
               PV := LIC_DRUM_PV, CSP := LIC_DRUM_CSP, STS := LIC_DRUM_STS);
      FIC_FW(PV_IN := fw, CSP_IN := fw, CSP_OK := TRUE, TRK := ficCas, TRK_VAL := LIC_DRUM.Q,
             DTS := dts, RESYNC := RT.RESYNC, PV_MIN := 0.0, PV_MAX := 2600.0, CAS_CFG := TRUE,
             SP := FIC_FW_SP, OUT := FIC_FW_OUT, MODE := FIC_FW_MODE, KP := FIC_FW_KP, TI := FIC_FW_TI, TD := FIC_FW_TD,
             PV := FIC_FW_PV, CSP := FIC_FW_CSP, STS := FIC_FW_STS);
    ELSE
      (* 3-element: level master trims the steam flow feed-forward, flow loop is the slave *)
      LIC_DRUM(PV_IN := lvl, TRK := NOT ficCas, TRK_VAL := e3Trk,
               DTS := dts, RESYNC := RT.RESYNC OR e3Changed, PV_MIN := -500.0, PV_MAX := 500.0,
               SP := LIC_DRUM_SP, OUT := LIC_DRUM_OUT, MODE := LIC_DRUM_MODE, KP := LIC_DRUM_KP, TI := LIC_DRUM_TI, TD := LIC_DRUM_TD,
               PV := LIC_DRUM_PV, CSP := LIC_DRUM_CSP, STS := LIC_DRUM_STS);
      FIC_FW(PV_IN := fw, CSP_IN := LIMIT(0.0, ff + (LIC_DRUM.Q - 50.0) * TRIM_GAIN, 2600.0), CSP_OK := TRUE, TRK := FALSE,
             DTS := dts, RESYNC := RT.RESYNC, PV_MIN := 0.0, PV_MAX := 2600.0, CAS_CFG := TRUE,
             SP := FIC_FW_SP, OUT := FIC_FW_OUT, MODE := FIC_FW_MODE, KP := FIC_FW_KP, TI := FIC_FW_TI, TD := FIC_FW_TD,
             PV := FIC_FW_PV, CSP := FIC_FW_CSP, STS := FIC_FW_STS);
    END_IF;
    Q_FCV_DMD := FIC_FW.Q;
    LVL_AUTO := LIC_DRUM.AUTO AND ficCas;

    (* ---- boiler feed pumps: standby start on a partner trip (latched until the operator's STOP) *)
    nRun := 0;
    IF I_BFP_A_RUN THEN nRun := nRun + 1; END_IF;
    IF I_BFP_B_RUN THEN nRun := nRun + 1; END_IF;
    IF I_BFP_C_RUN THEN nRun := nRun + 1; END_IF;
    BFP_RUNNING := nRun;
    daLvl := I_DA_LVL;
    tripA := I_BFP_A_TRIP OR (BFP_A.LATCHED AND NOT init);
    tripB := I_BFP_B_TRIP OR (BFP_B.LATCHED AND NOT init);
    tripC := I_BFP_C_TRIP OR (BFP_C.LATCHED AND NOT init);
    BFP_A(RUN_FB := I_BFP_A_RUN, TRIP_FB := I_BFP_A_TRIP, PERMIT := daLvl > 1200.0 AND SC_BFPA_OUT <= 10.0,
          AUTO_START := (tripB OR tripC) AND nRun < 3, SYNC := init,
          START := BFP_A_START, STOP := BFP_A_STOP, MODE := BFP_A_MODE, CMD := Q_BFP_A_CMD,
          RUN := BFP_A_RUN, TRIP := BFP_A_TRIP, PERM := BFP_A_PERM, ILK_T := BFP_A_ILK);
    IF I_BFP_A_RUN AND NOT runPrevA AND BFP_A.IS_AUTO AND (tripB OR tripC) THEN joinA := TRUE; END_IF;
    runPrevA := I_BFP_A_RUN;
    tripA := I_BFP_A_TRIP OR BFP_A.LATCHED;
    BFP_B(RUN_FB := I_BFP_B_RUN, TRIP_FB := I_BFP_B_TRIP, PERMIT := daLvl > 1200.0 AND SC_BFPB_OUT <= 10.0,
          AUTO_START := (tripA OR tripC) AND nRun < 3, SYNC := init,
          START := BFP_B_START, STOP := BFP_B_STOP, MODE := BFP_B_MODE, CMD := Q_BFP_B_CMD,
          RUN := BFP_B_RUN, TRIP := BFP_B_TRIP, PERM := BFP_B_PERM, ILK_T := BFP_B_ILK);
    IF I_BFP_B_RUN AND NOT runPrevB AND BFP_B.IS_AUTO AND (tripA OR tripC) THEN joinB := TRUE; END_IF;
    runPrevB := I_BFP_B_RUN;
    tripB := I_BFP_B_TRIP OR BFP_B.LATCHED;
    BFP_C(RUN_FB := I_BFP_C_RUN, TRIP_FB := I_BFP_C_TRIP, PERMIT := daLvl > 1200.0 AND SC_BFPC_OUT <= 10.0,
          AUTO_START := (tripA OR tripB) AND nRun < 3, SYNC := init,
          START := BFP_C_START, STOP := BFP_C_STOP, MODE := BFP_C_MODE, CMD := Q_BFP_C_CMD,
          RUN := BFP_C_RUN, TRIP := BFP_C_TRIP, PERM := BFP_C_PERM, ILK_T := BFP_C_ILK);
    IF I_BFP_C_RUN AND NOT runPrevC AND BFP_C.IS_AUTO AND (tripA OR tripB) THEN joinC := TRUE; END_IF;
    runPrevC := I_BFP_C_RUN;

    (* ---- BFP master: feedwater valve differential pressure *)
    dp := I_FW_HDR_PRESS - I_DRUM_PRESS;
    FW_DP := dp;
    anyAuto := (I_BFP_A_RUN AND SC_BFPA_MODE = 1) OR (I_BFP_B_RUN AND SC_BFPB_MODE = 1) OR (I_BFP_C_RUN AND SC_BFPC_MODE = 1);
    avgScoop := 0.0;
    IF I_BFP_A_RUN THEN avgScoop := avgScoop + SC_BFPA_OUT; END_IF;
    IF I_BFP_B_RUN THEN avgScoop := avgScoop + SC_BFPB_OUT; END_IF;
    IF I_BFP_C_RUN THEN avgScoop := avgScoop + SC_BFPC_OUT; END_IF;
    IF nRun > 0 THEN avgScoop := avgScoop / DINT_TO_REAL(nRun); END_IF;
    (* DP setpoint program: 10 bar at no load, 12 bar at 30 %, 20 bar at 100 % steam flow *)
    IF steamPct <= 30.0 THEN
      dpSp := 10.0 + LIMIT(0.0, steamPct, 30.0) / 30.0 * 2.0;
    ELSE
      dpSp := 12.0 + (MIN(steamPct, 100.0) - 30.0) / 70.0 * 8.0;
    END_IF;
    PIC_FWDP(PV_IN := dp, CSP_IN := dpSp, CSP_OK := DP_SP_MODE = 1, TRK := nRun = 0 OR NOT anyAuto, TRK_VAL := avgScoop,
             DTS := dts, RESYNC := RT.RESYNC, PV_MIN := 0.0, PV_MAX := 50.0, CAS_CFG := TRUE,
             SP := PIC_FWDP_SP, OUT := PIC_FWDP_OUT, MODE := PIC_FWDP_MODE, KP := PIC_FWDP_KP, TI := PIC_FWDP_TI, TD := PIC_FWDP_TD,
             PV := PIC_FWDP_PV, CSP := PIC_FWDP_CSP, STS := PIC_FWDP_STS);
    master := PIC_FWDP.Q;
    BFP_MASTER := master;
    SC_BFPA(AUTO_IN := master, FB_IN := LIMIT(0.0, (I_BFP_A_SPEED - 1500.0) / 39.0, 100.0), FORCE_MAN := NOT I_BFP_A_RUN,
            TRK := NOT I_BFP_A_RUN, TRK_VAL := 0.0, RATE := 3.0, DTS := dts, INIT := init, INIT_KEEP := keep, JOIN := joinA,
            OUT := SC_BFPA_OUT, MODE := SC_BFPA_MODE, BIAS := SC_BFPA_BIAS, IN_TAG := SC_BFPA_IN, FB_TAG := SC_BFPA_FB, STS := SC_BFPA_STS);
    SC_BFPB(AUTO_IN := master, FB_IN := LIMIT(0.0, (I_BFP_B_SPEED - 1500.0) / 39.0, 100.0), FORCE_MAN := NOT I_BFP_B_RUN,
            TRK := NOT I_BFP_B_RUN, TRK_VAL := 0.0, RATE := 3.0, DTS := dts, INIT := init, INIT_KEEP := keep, JOIN := joinB,
            OUT := SC_BFPB_OUT, MODE := SC_BFPB_MODE, BIAS := SC_BFPB_BIAS, IN_TAG := SC_BFPB_IN, FB_TAG := SC_BFPB_FB, STS := SC_BFPB_STS);
    SC_BFPC(AUTO_IN := master, FB_IN := LIMIT(0.0, (I_BFP_C_SPEED - 1500.0) / 39.0, 100.0), FORCE_MAN := NOT I_BFP_C_RUN,
            TRK := NOT I_BFP_C_RUN, TRK_VAL := 0.0, RATE := 3.0, DTS := dts, INIT := init, INIT_KEEP := keep, JOIN := joinC,
            OUT := SC_BFPC_OUT, MODE := SC_BFPC_MODE, BIAS := SC_BFPC_BIAS, IN_TAG := SC_BFPC_IN, FB_TAG := SC_BFPC_FB, STS := SC_BFPC_STS);
    joinA := FALSE; joinB := FALSE; joinC := FALSE;
    Q_BFP_A_SPD_DMD := SC_BFPA.Q;
    Q_BFP_B_SPD_DMD := SC_BFPB.Q;
    Q_BFP_C_SPD_DMD := SC_BFPC.Q;
    (* runback only if the standby pump has not restored two running pumps within 10 s *)
    T_RBBFP(IN := nRun < 2 AND steamPct > 58.0 AND I_GCB_CLOSED, PT := 10.0, DTS := dts, INIT := init);
    RB_BFP := T_RBBFP.Q;

    (* ---- deaerator level and pressure *)
    cep := I_CEP_A_RUN OR I_CEP_B_RUN;
    LIC_DA(PV_IN := daLvl, TRK := NOT cep, TRK_VAL := 0.0,
           DTS := dts, RESYNC := RT.RESYNC, PV_MIN := 0.0, PV_MAX := 3000.0,
           SP := LIC_DA_SP, OUT := LIC_DA_OUT, MODE := LIC_DA_MODE, KP := LIC_DA_KP, TI := LIC_DA_TI, TD := LIC_DA_TD,
           PV := LIC_DA_PV, CSP := LIC_DA_CSP, STS := LIC_DA_STS);
    Q_DA_CV_DMD := LIC_DA.Q;
    PIC_DA(PV_IN := I_DA_PRESS,
           DTS := dts, RESYNC := RT.RESYNC, PV_MIN := 0.0, PV_MAX := 10.0,
           SP := PIC_DA_SP, OUT := PIC_DA_OUT, MODE := PIC_DA_MODE, KP := PIC_DA_KP, TI := PIC_DA_TI, TD := PIC_DA_TD,
           PV := PIC_DA_PV, CSP := PIC_DA_CSP, STS := PIC_DA_STS);
    Q_PEG_DMD := PIC_DA.Q;

    (* ---- blowdown and HP heaters *)
    EBD(OPENED_FB := I_EBD_OPEN, AUTO_OPEN := lvl > 150.0, AUTO_CLOSE := lvl < 50.0, SYNC := init,
        OPEN := EBD_OPEN, CLOSE := EBD_CLOSE, MODE := EBD_MODE, CMD := Q_EBD_CMD,
        OPENED := EBD_OPENED, CLOSED := EBD_CLOSED, PERM := EBD_PERM, ILK := EBD_ILK);
    HPH(OPENED_FB := I_HPH_IN_SERVICE, SYNC := init,
        OPEN := HPH_OPEN, CLOSE := HPH_CLOSE, MODE := HPH_MODE, CMD := Q_HPH_CMD,
        OPENED := HPH_OPENED, CLOSED := HPH_CLOSED, PERM := HPH_PERM, ILK := HPH_ILK);
    HIC_CBD(AUTO_IN := 0.0, FB_IN := I_CBD_FB, DTS := dts, INIT := init, INIT_KEEP := keepCbd,
            OUT := HIC_CBD_OUT, MODE := HIC_CBD_MODE, BIAS := HIC_CBD_BIAS, IN_TAG := HIC_CBD_IN, FB_TAG := HIC_CBD_FB, STS := HIC_CBD_STS);
    Q_CBD_DMD := HIC_CBD.Q;
  END_IF;
END_PROGRAM

(* ---- GEN.st ---- *)
(* GEN - Generator, Excitation & Synchronising
   Generator protection with lockout relay 86G (first-out cause), field breaker (41) and
   generator breaker (52G), automatic synchroniser (speed matching via DEH, voltage matching
   via the AVR, advance-angle closing), AVR with MVAr / power-factor control and over / under
   excitation limiters, field forcing to no-load excitation on load rejection.
   Naming: I_* field inputs, Q_* field outputs, P_<PEER>_* peer status, W_<PEER>_* writes to
   a peer, IO_* bridge signals. *)
PROGRAM GEN_MAIN
(*@IO*)
  VAR
    RT : FB_PLC_RUNTIME;
    FCB : FB_ONOFF;
    GCB : FB_ONOFF;
    AVR : FB_LOOP;
    T_OOS : FB_TONS;           (* loss of field / pole slip *)
    T_REVP : FB_TONS;          (* reverse power *)
    T_OV : FB_TONS;            (* overvoltage *)
    T_FREQ : FB_TONS;          (* over / under frequency *)
    T_VHZ : FB_TONS;           (* over-excitation V/Hz *)
    T_OC : FB_TONS;            (* overcurrent *)
    T_LFP : FB_TONS;           (* low forward power after turbine trip *)
    dts : REAL;
    init : BOOL;
    speed : REAL;
    freq : REAL;
    vPu : REAL;
    gPu : REAL;
    vhzV : REAL;
    gcbIn : BOOL;
    fcbIn : BOOL;
    mw : REAL;
    slip : REAL;
    phase : REAL;
    ifPu : REAL;
    dV : REAL;
    dehOk : BOOL;
    dehLatched : BOOL;
    dehTripped : BOOL;
    dehSpeedMode : BOOL;
    c : ARRAY[1..10] OF BOOL;  (* protection functions, by trip cause number *)
    firstOut : DINT;
    lock : BOOL;
    cause : DINT;
    faultActive : BOOL;
    syncCheck : BOOL;
    syncPerm : BOOL;
    sync : DINT;               (* 0 OFF, 1 WAIT, 2 MATCH, 3 CLOSING, 4 DONE *)
    syncT : REAL;
    autoClose : BOOL;
    adj : REAL;
    vTarget : REAL;
    advance : REAL;
    qTarget : REAL;
    qErr : REAL;
    oel : BOOL;
    uel : BOOL;
    gcbPrev : BOOL;
    gcbOpened : BOOL;
    excHi : REAL;
    excLo : REAL;
  END_VAR
  VAR CONSTANT
    SLIP_TARGET : REAL := 0.08;   (* Hz, generator slightly faster than the grid *)
    RATED_KA : REAL := 21.6;       (* kA *)
  END_VAR

  (* ---------------------------------------------------------------- runtime services *)
  RT(SIM_MS := I_SIM_TIME_MS, IC_SEQ := IO_IC_SEQ, IC_ID := IO_IC_ID, IC_SNAP := IO_IC_SNAP, CYCLE_MS := 50.0,
     HEARTBEAT := HEARTBEAT, SCAN_COUNT := SCAN_COUNT, SCAN_MS := SCAN_MS, SIM_DT := SIM_DT,
     IC_APPLIED := IC_APPLIED, IC_ACK := IC_ACK);
  dts := RT.DTS;
  init := RT.IC_INIT;
  HEALTHY := IO_COMM_PLANT AND RT.READY;
  COMM_PLANT := IO_COMM_PLANT OR NOT RT.READY;   (* not reported before the bridge has initialised the PLC *)
  COMM_DEH := IO_COMM_DEH OR RT.GRACE OR NOT RT.READY;

  IF init THEN
    lock := FALSE;
    cause := 0;
    sync := 0;
    syncT := 0.0;
    gcbPrev := FALSE;
  END_IF;

  (* ---------------------------------------------------------------- built-in initial condition *)
  IF RT.IC_BUILTIN THEN
    IF I_FCB_CLOSED THEN
      AVR_OUT := I_FIELD_AMPS / 2400.0;
      AVR_SP := I_GEN_KV;
      AVR_MODE := 1;
    ELSE
      AVR_OUT := 0.0;
      AVR_SP := 22.0;
      AVR_MODE := 0;
    END_IF;
    FCB_MODE := 0;
    GCB_MODE := 0;
  END_IF;

  IF RT.READY THEN
    speed := I_SPEED_B;
    freq := MAX(1.0, speed / 60.0);
    vPu := I_GEN_KV / 22.0;
    gPu := I_GRID_KV / 400.0;
    vhzV := vPu / (freq / 60.0);
    gcbIn := I_GCB_CLOSED;
    fcbIn := I_FCB_CLOSED;
    mw := I_GEN_MW;
    slip := I_SYNC_SLIP;
    phase := I_SYNC_PHASE;
    ifPu := I_FIELD_AMPS / 2400.0;
    dehOk := IO_COMM_DEH;
    dehLatched := dehOk AND P_DEH_LATCHED;
    IF dehOk THEN dehTripped := P_DEH_TRIPPED; ELSE dehTripped := TRUE; END_IF;
    dehSpeedMode := dehOk AND P_DEH_MODE = 1;
    V_PU := vPu;
    GRID_V_PU := gPu;
    VHZ := vhzV;
    dV := (vPu - gPu) * 100.0;
    DV_PCT := dV;

    (* ---------------------------------------------------------------- protection (86G lockout) *)
    T_OOS(IN := gcbIn AND (I_OUT_OF_STEP OR ifPu < 0.15), PT := 0.5, DTS := dts, INIT := init);
    IF dehTripped THEN
      T_REVP(IN := gcbIn AND mw < -4.0, PT := 2.0, DTS := dts, INIT := init);
    ELSE
      T_REVP(IN := gcbIn AND mw < -4.0, PT := 5.0, DTS := dts, INIT := init);
    END_IF;
    T_OV(IN := fcbIn AND vPu > 1.18, PT := 5.0, DTS := dts, INIT := init);
    T_FREQ(IN := gcbIn AND (freq < 57.5 OR freq > 61.8), PT := 5.0, DTS := dts, INIT := init);
    T_VHZ(IN := fcbIn AND vhzV > 1.12, PT := 5.0, DTS := dts, INIT := init);
    T_OC(IN := I_GEN_KA > 1.3 * RATED_KA, PT := 10.0, DTS := dts, INIT := init);
    T_LFP(IN := dehTripped AND gcbIn AND mw < 10.0, PT := 20.0, DTS := dts, INIT := init);
    c[1] := TRIP_86;                       (* manual trip *)
    c[2] := I_GEN_DIFF_RELAY;              (* 87G *)
    c[3] := T_OOS.Q;                       (* 40 / 78 *)
    c[4] := T_REVP.Q;                      (* 32 *)
    c[5] := T_OV.Q OR vPu > 1.4;           (* 59, instantaneous above 1.4 pu *)
    c[6] := T_FREQ.Q;                      (* 81 *)
    c[7] := T_VHZ.Q;                       (* 24 *)
    c[8] := I_STATOR_TEMP > 125.0;
    c[9] := T_OC.Q;                        (* 51 *)
    c[10] := T_LFP.Q;                      (* sequential tripping *)
    REV_POWER := gcbIn AND mw < -2.0;
    firstOut := FIRST_OUT(C1 := c[1], C2 := c[2], C3 := c[3], C4 := c[4], C5 := c[5], C6 := c[6], C7 := c[7], C8 := c[8], C9 := c[9],
                          C10 := c[10]);
    IF NOT lock AND firstOut > 0 THEN
      lock := TRUE;
      cause := firstOut;
      sync := 0;
    END_IF;
    IF RESET_86 THEN
      faultActive := c[2] OR c[3] OR c[5] OR c[7] OR c[8];
      IF lock AND NOT faultActive THEN
        lock := FALSE;
        cause := 0;
      END_IF;
    END_IF;

    (* ---------------------------------------------------------------- breakers *)
    syncCheck := NOT gcbIn AND fcbIn AND ABS(slip) < 0.2 AND ABS(phase) < 15.0 AND ABS(dV) < 5.0;
    SYNC_CHECK := syncCheck;
    FCB(OPENED_FB := fcbIn, PERMIT := speed > 3420.0 AND NOT lock AND dehLatched, ILK_CLOSE := lock OR speed < 3000.0,
        RESET_ON_LOSS := TRUE, SYNC := init,
        OPEN := FCB_OPEN, CLOSE := FCB_CLOSE, MODE := FCB_MODE, CMD := Q_FCB_CMD,
        OPENED := FCB_OPENED, CLOSED := FCB_CLOSED, PERM := FCB_PERM, ILK := FCB_ILK);

    (* ---------------------------------------------------------------- auto synchroniser *)
    autoClose := FALSE;
    adj := 0.0;
    IF SYNC_ON AND NOT gcbIn THEN sync := 1; END_IF;
    IF SYNC_OFF THEN sync := 0; END_IF;
    syncPerm := dehLatched AND dehSpeedMode AND speed > 3540.0 AND fcbIn AND AVR_MODE <> 0 AND NOT lock AND NOT gcbIn;
    CASE sync OF
      1: (* waiting for permissives *)
        IF syncPerm THEN sync := 2; END_IF;
      2: (* matching speed and voltage *)
        IF NOT syncPerm THEN
          sync := 1;
        ELSE
          adj := LIMIT(-4.0, (SLIP_TARGET - slip) * 60.0 * 0.6, 4.0);
          vTarget := gPu * 22.0 * 1.005;
          AVR_SP := AVR_SP + LIMIT(-0.2 * dts, vTarget - AVR_SP, 0.2 * dts);
          advance := 360.0 * slip * 0.08;   (* breaker closing time 80 ms *)
          IF slip > 0.02 AND slip < 0.2 AND ABS(dV) < 2.0 AND phase < -advance + 4.0 AND phase > -advance - 6.0 THEN
            autoClose := TRUE;
            sync := 3;
            syncT := 0.0;
          END_IF;
        END_IF;
      3: (* closing *)
        autoClose := TRUE;
        syncT := syncT + dts;
        IF gcbIn THEN
          sync := 4;
          syncT := 0.0;
        ELSIF syncT > 2.0 THEN
          sync := 2;
        END_IF;
      4: (* synchronised *)
        syncT := syncT + dts;
        IF syncT > 5.0 THEN sync := 0; END_IF;
    END_CASE;
    IF gcbIn AND sync <> 4 AND sync <> 0 THEN sync := 4; END_IF;
    SYNC_STATE := sync;
    W_DEH_SYNC_ADJ := adj;
    IF sync = 2 OR sync = 3 THEN W_DEH_SYNC_ACTIVE := 1; ELSE W_DEH_SYNC_ACTIVE := 0; END_IF;

    GCB(OPENED_FB := gcbIn, PERMIT := (syncCheck OR gcbIn) AND NOT lock AND dehLatched, ILK_CLOSE := lock,
        RESET_ON_LOSS := TRUE, CMD_SET := autoClose, CMD_VAL := TRUE, SYNC := init,
        OPEN := GCB_OPEN, CLOSE := GCB_CLOSE, MODE := GCB_MODE, CMD := Q_GCB_CMD,
        OPENED := GCB_OPENED, CLOSED := GCB_CLOSED, PERM := GCB_PERM, ILK := GCB_ILK);

    (* ---------------------------------------------------------------- AVR & limiters *)
    (* on line: MVAr or power-factor control trims the voltage setpoint slowly *)
    IF gcbIn AND AVR_MODE <> 0 AND EXC_MODE > 0 THEN
      IF EXC_MODE = 1 THEN
        qTarget := MVAR_SP;
      ELSE
        qTarget := mw * TAN(ACOS(LIMIT(0.7, PF_SP, 1.0)));
      END_IF;
      qErr := qTarget - I_GEN_MVAR;
      AVR_SP := LIMIT(20.0, AVR_SP + LIMIT(-1.0, qErr / 300.0, 1.0) * 0.05 * dts, 24.2);
    END_IF;
    (* off line: V/Hz limiter *)
    IF NOT gcbIn AND AVR_MODE <> 0 THEN
      AVR_SP := MIN(AVR_SP, 22.0 * 1.05 * (freq / 60.0));
    END_IF;
    oel := ifPu > 2.1;
    uel := gcbIn AND I_GEN_MVAR < -0.3 * MAX(0.0, mw) - 120.0;
    OEL_ACTIVE := oel;
    UEL_ACTIVE := uel;
    (* load rejection: force the field down to no-load excitation so the voltage stays near rated *)
    gcbOpened := NOT gcbIn AND gcbPrev;
    gcbPrev := gcbIn;
    IF gcbOpened AND AVR_MODE <> 0 THEN
      AVR_OUT := 1.0;
      AVR_SP := 22.0;
      AVR_MODE := 1;
      EXC_MODE := 0;
    END_IF;
    IF oel THEN excHi := ifPu; ELSE excHi := 2.3; END_IF;
    IF uel THEN excLo := ifPu + 0.005; ELSE excLo := 0.0; END_IF;
    AVR(PV_IN := I_GEN_KV, TRK := NOT fcbIn, TRK_VAL := 0.0, OUT_HI := excHi, OUT_LO := excLo,
        DTS := dts, RESYNC := RT.RESYNC OR gcbOpened, PV_MIN := 0.0, PV_MAX := 30.0, OUT_MIN := 0.0, OUT_MAX := 2.3,
        SP_TRACK := FALSE, REF_DT := 0.15,
        SP := AVR_SP, OUT := AVR_OUT, MODE := AVR_MODE, KP := AVR_KP, TI := AVR_TI, TD := AVR_TD,
        PV := AVR_PV, CSP := AVR_CSP, STS := AVR_STS);
    Q_EXC_DMD := AVR.Q;

    LOCKOUT_86 := lock;
    TRIP_CAUSE := cause;
  END_IF;

  (* operator pulses are consumed in the scan they arrive *)
  SYNC_ON := FALSE;
  SYNC_OFF := FALSE;
  RESET_86 := FALSE;
  TRIP_86 := FALSE;
END_PROGRAM
